// TIA Portal V20 program export: 0 tag tables, 53 data types, 23 data blocks, 177 code blocks (in call order from the OBs), 3 instance data blocks

TYPE "FRK_Access"
// stored: IsFailsafeCompliant false
   STRUCT
      CurrentLevel : DInt;
      CurrentUser : String[32];
      LoginFailed : Bool;
      Policy { S7_SetPoint := 'True'} : "ST_AccessPolicy";
      SessionGeneration : UDInt;
      LoginBusy : Bool;
      LoginResultSequence : UDInt;
      LoginTimeoutMs : UDInt;
      PolicySlot { ExternalAccessible := 'False'; ExternalVisible := 'False'; ExternalWritable := 'False'} : Int;
      PolicyLost { ExternalAccessible := 'False'; ExternalVisible := 'False'; ExternalWritable := 'False'} : Bool;
      PolicyLossAlarm { ExternalAccessible := 'False'; ExternalVisible := 'False'; ExternalWritable := 'False'} : Int;
      UserLossAlarm { ExternalAccessible := 'False'; ExternalVisible := 'False'; ExternalWritable := 'False'} : Int;
      ProviderGeneration { ExternalAccessible := 'False'; ExternalVisible := 'False'; ExternalWritable := 'False'} : UDInt;
      CandidateGeneration { ExternalAccessible := 'False'; ExternalVisible := 'False'; ExternalWritable := 'False'} : UDInt;
      ProviderEnabled { ExternalAccessible := 'False'; ExternalVisible := 'False'; ExternalWritable := 'False'} : Bool;
      LastActivity { ExternalAccessible := 'False'; ExternalVisible := 'False'; ExternalWritable := 'False'} : UDInt;
      LoginSince { ExternalAccessible := 'False'; ExternalVisible := 'False'; ExternalWritable := 'False'} : UDInt;
      LoginSequence { ExternalAccessible := 'False'; ExternalVisible := 'False'; ExternalWritable := 'False'} : UDInt;
      CandidateUser { ExternalAccessible := 'False'; ExternalVisible := 'False'; ExternalWritable := 'False'} : String[32];
      CandidateLevel { ExternalAccessible := 'False'; ExternalVisible := 'False'; ExternalWritable := 'False'} : DInt;
      Round { ExternalAccessible := 'False'; ExternalVisible := 'False'; ExternalWritable := 'False'} : DInt;
      Salt { ExternalAccessible := 'False'; ExternalVisible := 'False'; ExternalWritable := 'False'} : Array[0..15] of Byte;
      Digest { ExternalAccessible := 'False'; ExternalVisible := 'False'; ExternalWritable := 'False'} : Array[0..31] of Byte;
      Expected { ExternalAccessible := 'False'; ExternalVisible := 'False'; ExternalWritable := 'False'} : Array[0..31] of Byte;
   END_STRUCT;
END_TYPE

TYPE "FRK_AccessPolicyImage"
// stored: IsFailsafeCompliant false
   STRUCT
      SchemaVersion { ExternalAccessible := 'False'; ExternalVisible := 'False'; ExternalWritable := 'False'} : UInt;
      Scope { ExternalAccessible := 'False'; ExternalVisible := 'False'; ExternalWritable := 'False'} : String[80];
      Generation { ExternalAccessible := 'False'; ExternalVisible := 'False'; ExternalWritable := 'False'} : UDInt;
      Policy { ExternalAccessible := 'False'; ExternalVisible := 'False'; ExternalWritable := 'False'; S7_SetPoint := 'True'} : "ST_AccessPolicy";
      Checksum { ExternalAccessible := 'False'; ExternalVisible := 'False'; ExternalWritable := 'False'} : DWord;
   END_STRUCT;
END_TYPE

TYPE "FRK_AlarmLog"
// stored: IsFailsafeCompliant false
   STRUCT
      Active { S7_SetPoint := 'True'} : Array[1..16] of "ST_AlarmEvent";
      NActive : Int;
      Ring { S7_SetPoint := 'True'} : Array[1..64] of "ST_AlarmEvent";
      RingHead : Int;
      Blocking : Bool;
      Truncated : Bool;
      ComeMs { ExternalAccessible := 'False'; ExternalVisible := 'False'; ExternalWritable := 'False'} : Array[1..16] of UDInt;
      Automatic { ExternalAccessible := 'False'; ExternalVisible := 'False'; ExternalWritable := 'False'} : Array[1..16] of Bool;
      Touched { ExternalAccessible := 'False'; ExternalVisible := 'False'; ExternalWritable := 'False'} : Array[1..16] of Bool;
      RingUsed { ExternalAccessible := 'False'; ExternalVisible := 'False'; ExternalWritable := 'False'} : Int;
      SinkEnabled { ExternalAccessible := 'False'; ExternalVisible := 'False'; ExternalWritable := 'False'} : Bool;
   END_STRUCT;
END_TYPE

TYPE "FRK_Carrier"
// stored: IsFailsafeCompliant false
   STRUCT
      Enabled { ExternalAccessible := 'False'; ExternalVisible := 'False'; ExternalWritable := 'False'} : Bool;
      Kind { ExternalAccessible := 'False'; ExternalVisible := 'False'; ExternalWritable := 'False'} : DInt;
      Serial { ExternalAccessible := 'False'; ExternalVisible := 'False'; ExternalWritable := 'False'} : UDInt;
      Context { ExternalAccessible := 'False'; ExternalVisible := 'False'; ExternalWritable := 'False'; S7_SetPoint := 'True'} : "ST_PartContext";
      Written { ExternalAccessible := 'False'; ExternalVisible := 'False'; ExternalWritable := 'False'; S7_SetPoint := 'True'} : "ST_PartContext";
      Writes { ExternalAccessible := 'False'; ExternalVisible := 'False'; ExternalWritable := 'False'} : UDInt;
   END_STRUCT;
END_TYPE

TYPE "FRK_ConfigCursor"
// stored: IsFailsafeCompliant false
   STRUCT
      Position { ExternalAccessible := 'False'; ExternalVisible := 'False'; ExternalWritable := 'False'} : DInt;
      First { ExternalAccessible := 'False'; ExternalVisible := 'False'; ExternalWritable := 'False'} : DInt;
   END_STRUCT;
END_TYPE

TYPE "FRK_ConfigSlot"
// stored: IsFailsafeCompliant false
   STRUCT
      SchemaVersion { ExternalAccessible := 'False'; ExternalVisible := 'False'; ExternalWritable := 'False'} : UInt;
      Used { ExternalAccessible := 'False'; ExternalVisible := 'False'; ExternalWritable := 'False'} : Bool;
      ModelCode { ExternalAccessible := 'False'; ExternalVisible := 'False'; ExternalWritable := 'False'} : String[64];
      Record { ExternalAccessible := 'False'; ExternalVisible := 'False'; ExternalWritable := 'False'; S7_SetPoint := 'True'} : "ST_ConfigRecord";
   END_STRUCT;
END_TYPE

TYPE "FRK_ConfigValue"
// stored: IsFailsafeCompliant false
   STRUCT
      Number { ExternalAccessible := 'False'; ExternalVisible := 'False'; ExternalWritable := 'False'} : LInt;
      Flag { ExternalAccessible := 'False'; ExternalVisible := 'False'; ExternalWritable := 'False'} : Bool;
      Text { ExternalAccessible := 'False'; ExternalVisible := 'False'; ExternalWritable := 'False'} : String[80];
   END_STRUCT;
END_TYPE

TYPE "FRK_Core"
// stored: IsFailsafeCompliant false
   STRUCT
      Named { ExternalAccessible := 'False'; ExternalVisible := 'False'; ExternalWritable := 'False'} : Bool;
      Initialized { ExternalAccessible := 'False'; ExternalVisible := 'False'; ExternalWritable := 'False'} : Bool;
      RegIndex { ExternalAccessible := 'False'; ExternalVisible := 'False'; ExternalWritable := 'False'} : DInt;
      ParentIndex { ExternalAccessible := 'False'; ExternalVisible := 'False'; ExternalWritable := 'False'} : DInt;
      ModuleType { ExternalAccessible := 'False'; ExternalVisible := 'False'; ExternalWritable := 'False'} : DInt;
      Exec { ExternalAccessible := 'False'; ExternalVisible := 'False'; ExternalWritable := 'False'} : DInt;
      ExecPrev { ExternalAccessible := 'False'; ExternalVisible := 'False'; ExternalWritable := 'False'} : Bool;
      AbortPrev { ExternalAccessible := 'False'; ExternalVisible := 'False'; ExternalWritable := 'False'} : Bool;
      Armed { ExternalAccessible := 'False'; ExternalVisible := 'False'; ExternalWritable := 'False'} : Bool;
      Command { ExternalAccessible := 'False'; ExternalVisible := 'False'; ExternalWritable := 'False'} : DInt;
      CommandLabel { ExternalAccessible := 'False'; ExternalVisible := 'False'; ExternalWritable := 'False'} : String[120];
      Dispatch { ExternalAccessible := 'False'; ExternalVisible := 'False'; ExternalWritable := 'False'} : Bool;
      EvInit { ExternalAccessible := 'False'; ExternalVisible := 'False'; ExternalWritable := 'False'} : Bool;
      EvCommandStart { ExternalAccessible := 'False'; ExternalVisible := 'False'; ExternalWritable := 'False'} : Bool;
      ReleasePending { ExternalAccessible := 'False'; ExternalVisible := 'False'; ExternalWritable := 'False'} : Bool;
      EvAbort { ExternalAccessible := 'False'; ExternalVisible := 'False'; ExternalWritable := 'False'} : Bool;
      EvAbortInError { ExternalAccessible := 'False'; ExternalVisible := 'False'; ExternalWritable := 'False'} : Bool;
      EvModeExit { ExternalAccessible := 'False'; ExternalVisible := 'False'; ExternalWritable := 'False'} : Bool;
      EvModeChanged { ExternalAccessible := 'False'; ExternalVisible := 'False'; ExternalWritable := 'False'} : Bool;
      "Step" { ExternalAccessible := 'False'; ExternalVisible := 'False'; ExternalWritable := 'False'} : DInt;
      HookResult { ExternalAccessible := 'False'; ExternalVisible := 'False'; ExternalWritable := 'False'} : DInt;
      Held { ExternalAccessible := 'False'; ExternalVisible := 'False'; ExternalWritable := 'False'} : Bool;
      HoldReq { ExternalAccessible := 'False'; ExternalVisible := 'False'; ExternalWritable := 'False'} : Bool;
      HoldReason { ExternalAccessible := 'False'; ExternalVisible := 'False'; ExternalWritable := 'False'} : DInt;
      DiagTouched { ExternalAccessible := 'False'; ExternalVisible := 'False'; ExternalWritable := 'False'} : Bool;
      TimingOpen { ExternalAccessible := 'False'; ExternalVisible := 'False'; ExternalWritable := 'False'} : Bool;
      StartMs { ExternalAccessible := 'False'; ExternalVisible := 'False'; ExternalWritable := 'False'} : UDInt;
      LastNowMs { ExternalAccessible := 'False'; ExternalVisible := 'False'; ExternalWritable := 'False'} : UDInt;
      DeltaMs { ExternalAccessible := 'False'; ExternalVisible := 'False'; ExternalWritable := 'False'} : UDInt;
      ActiveMs { ExternalAccessible := 'False'; ExternalVisible := 'False'; ExternalWritable := 'False'} : UDInt;
      TimeoutMs { ExternalAccessible := 'False'; ExternalVisible := 'False'; ExternalWritable := 'False'} : UDInt;
      Timing { ExternalAccessible := 'False'; ExternalVisible := 'False'; ExternalWritable := 'False'; S7_SetPoint := 'True'} : "ST_ModuleTiming";
      FaultSlot { ExternalAccessible := 'False'; ExternalVisible := 'False'; ExternalWritable := 'False'} : Int;
      FaultHandled { ExternalAccessible := 'False'; ExternalVisible := 'False'; ExternalWritable := 'False'} : Bool;
   END_STRUCT;
END_TYPE

TYPE "FRK_DecisionSlot"
// stored: IsFailsafeCompliant false
   STRUCT
      RootIndex { ExternalAccessible := 'False'; ExternalVisible := 'False'; ExternalWritable := 'False'} : DInt;
      Owner { ExternalAccessible := 'False'; ExternalVisible := 'False'; ExternalWritable := 'False'} : DInt;
      Request { ExternalAccessible := 'False'; ExternalVisible := 'False'; ExternalWritable := 'False'; S7_SetPoint := 'True'} : "ST_DecisionRequest";
      Answer { ExternalAccessible := 'False'; ExternalVisible := 'False'; ExternalWritable := 'False'} : Int;
      AskedAt { ExternalAccessible := 'False'; ExternalVisible := 'False'; ExternalWritable := 'False'} : UDInt;
      OverlapLogged { ExternalAccessible := 'False'; ExternalVisible := 'False'; ExternalWritable := 'False'} : Bool;
      ResolutionLogged { ExternalAccessible := 'False'; ExternalVisible := 'False'; ExternalWritable := 'False'} : Bool;
   END_STRUCT;
END_TYPE

TYPE "FRK_JsonField"
// stored: IsFailsafeCompliant false
   STRUCT
      Key { ExternalAccessible := 'False'; ExternalVisible := 'False'; ExternalWritable := 'False'} : String[16];
      Text { ExternalAccessible := 'False'; ExternalVisible := 'False'; ExternalWritable := 'False'} : WString[160];
      Quoted { ExternalAccessible := 'False'; ExternalVisible := 'False'; ExternalWritable := 'False'} : Bool;
   END_STRUCT;
END_TYPE

TYPE "FRK_ManualConditionRow"
// stored: IsFailsafeCompliant false
   STRUCT
      Used { ExternalAccessible := 'False'; ExternalVisible := 'False'; ExternalWritable := 'False'} : Bool;
      Value { ExternalAccessible := 'False'; ExternalVisible := 'False'; ExternalWritable := 'False'} : DInt;
      Ok { ExternalAccessible := 'False'; ExternalVisible := 'False'; ExternalWritable := 'False'} : Bool;
      Diag { ExternalAccessible := 'False'; ExternalVisible := 'False'; ExternalWritable := 'False'; S7_SetPoint := 'True'} : "ST_Diagnostic";
      Bypassable { ExternalAccessible := 'False'; ExternalVisible := 'False'; ExternalWritable := 'False'} : Bool;
   END_STRUCT;
END_TYPE

TYPE "FRK_RegistryRow"
// stored: IsFailsafeCompliant false
   STRUCT
      Valid { ExternalAccessible := 'False'; ExternalVisible := 'False'; ExternalWritable := 'False'} : Bool;
      Parent { ExternalAccessible := 'False'; ExternalVisible := 'False'; ExternalWritable := 'False'} : DInt;
      ModuleType { ExternalAccessible := 'False'; ExternalVisible := 'False'; ExternalWritable := 'False'} : DInt;
      TypeId { ExternalAccessible := 'False'; ExternalVisible := 'False'; ExternalWritable := 'False'} : DInt;
      Capabilities { ExternalAccessible := 'False'; ExternalVisible := 'False'; ExternalWritable := 'False'} : DWord;
      Exec { ExternalAccessible := 'False'; ExternalVisible := 'False'; ExternalWritable := 'False'} : DInt;
      ReasonCode { ExternalAccessible := 'False'; ExternalVisible := 'False'; ExternalWritable := 'False'} : DInt;
      Severity { ExternalAccessible := 'False'; ExternalVisible := 'False'; ExternalWritable := 'False'} : DInt;
      AlarmBlocking { ExternalAccessible := 'False'; ExternalVisible := 'False'; ExternalWritable := 'False'} : Bool;
   END_STRUCT;
END_TYPE

TYPE "FRK_SetPayload"
// stored: IsFailsafeCompliant false
   STRUCT
      Info { ExternalAccessible := 'False'; ExternalVisible := 'False'; ExternalWritable := 'False'; S7_SetPoint := 'True'} : "ST_ConfigSetInfo";
      Records { ExternalAccessible := 'False'; ExternalVisible := 'False'; ExternalWritable := 'False'; S7_SetPoint := 'True'} : Array[1..24] of "ST_ConfigRecord";
   END_STRUCT;
END_TYPE

TYPE "FRK_SetWorkspace"
// stored: IsFailsafeCompliant false
   STRUCT
      Payload { ExternalAccessible := 'False'; ExternalVisible := 'False'; ExternalWritable := 'False'; S7_SetPoint := 'True'} : "FRK_SetPayload";
      Seen { ExternalAccessible := 'False'; ExternalVisible := 'False'; ExternalWritable := 'False'} : Array[1..24] of Bool;
      Matched { ExternalAccessible := 'False'; ExternalVisible := 'False'; ExternalWritable := 'False'} : Int;
      RejectScope { ExternalAccessible := 'False'; ExternalVisible := 'False'; ExternalWritable := 'False'} : String[80];
      RejectKey { ExternalAccessible := 'False'; ExternalVisible := 'False'; ExternalWritable := 'False'} : String[160];
      Importing { ExternalAccessible := 'False'; ExternalVisible := 'False'; ExternalWritable := 'False'} : Bool;
      Exporting { ExternalAccessible := 'False'; ExternalVisible := 'False'; ExternalWritable := 'False'} : Bool;
      NextLine { ExternalAccessible := 'False'; ExternalVisible := 'False'; ExternalWritable := 'False'} : Int;
      Generation { ExternalAccessible := 'False'; ExternalVisible := 'False'; ExternalWritable := 'False'} : UDInt;
      Received { ExternalAccessible := 'False'; ExternalVisible := 'False'; ExternalWritable := 'False'} : Int;
      Piece { ExternalAccessible := 'False'; ExternalVisible := 'False'; ExternalWritable := 'False'} : WString[480];
      Line { ExternalAccessible := 'False'; ExternalVisible := 'False'; ExternalWritable := 'False'} : WString[480];
      Fields { ExternalAccessible := 'False'; ExternalVisible := 'False'; ExternalWritable := 'False'; S7_SetPoint := 'True'} : Array[1..9] of "FRK_JsonField";
      FieldCount { ExternalAccessible := 'False'; ExternalVisible := 'False'; ExternalWritable := 'False'} : Int;
   END_STRUCT;
END_TYPE

TYPE "FRK_Unit"
// stored: IsFailsafeCompliant false
   STRUCT
      Initialized { ExternalAccessible := 'False'; ExternalVisible := 'False'; ExternalWritable := 'False'} : Bool;
      Mode { ExternalAccessible := 'False'; ExternalVisible := 'False'; ExternalWritable := 'False'} : DInt;
      RequestedMode { ExternalAccessible := 'False'; ExternalVisible := 'False'; ExternalWritable := 'False'} : DInt;
      ModePending { ExternalAccessible := 'False'; ExternalVisible := 'False'; ExternalWritable := 'False'} : Bool;
      ExitFirst { ExternalAccessible := 'False'; ExternalVisible := 'False'; ExternalWritable := 'False'} : Bool;
      RunReq { ExternalAccessible := 'False'; ExternalVisible := 'False'; ExternalWritable := 'False'} : Bool;
      AbortReq { ExternalAccessible := 'False'; ExternalVisible := 'False'; ExternalWritable := 'False'} : Bool;
      StopReq { ExternalAccessible := 'False'; ExternalVisible := 'False'; ExternalWritable := 'False'} : Bool;
      ModeSince { ExternalAccessible := 'False'; ExternalVisible := 'False'; ExternalWritable := 'False'} : UDInt;
      ReleaseChildren { ExternalAccessible := 'False'; ExternalVisible := 'False'; ExternalWritable := 'False'} : Bool;
      Clearing { ExternalAccessible := 'False'; ExternalVisible := 'False'; ExternalWritable := 'False'} : Bool;
      FaultLatched { ExternalAccessible := 'False'; ExternalVisible := 'False'; ExternalWritable := 'False'} : Bool;
      PrevError { ExternalAccessible := 'False'; ExternalVisible := 'False'; ExternalWritable := 'False'} : Bool;
      EvReset { ExternalAccessible := 'False'; ExternalVisible := 'False'; ExternalWritable := 'False'} : Bool;
      SeenSequence { ExternalAccessible := 'False'; ExternalVisible := 'False'; ExternalWritable := 'False'} : UDInt;
      RequestPending { ExternalAccessible := 'False'; ExternalVisible := 'False'; ExternalWritable := 'False'} : Bool;
      Request { ExternalAccessible := 'False'; ExternalVisible := 'False'; ExternalWritable := 'False'; S7_SetPoint := 'True'} : "ST_HmiRequest";
      RequestUser { ExternalAccessible := 'False'; ExternalVisible := 'False'; ExternalWritable := 'False'} : String[32];
      Permit { ExternalAccessible := 'False'; ExternalVisible := 'False'; ExternalWritable := 'False'} : Bool;
      PermitDiag { ExternalAccessible := 'False'; ExternalVisible := 'False'; ExternalWritable := 'False'; S7_SetPoint := 'True'} : "ST_Diagnostic";
      CarrierIndex { ExternalAccessible := 'False'; ExternalVisible := 'False'; ExternalWritable := 'False'} : DInt;
      Good { ExternalAccessible := 'False'; ExternalVisible := 'False'; ExternalWritable := 'False'} : UDInt;
      Nok { ExternalAccessible := 'False'; ExternalVisible := 'False'; ExternalWritable := 'False'} : UDInt;
      Rework { ExternalAccessible := 'False'; ExternalVisible := 'False'; ExternalWritable := 'False'} : UDInt;
      NokReason { ExternalAccessible := 'False'; ExternalVisible := 'False'; ExternalWritable := 'False'} : DInt;
      CascadePending { ExternalAccessible := 'False'; ExternalVisible := 'False'; ExternalWritable := 'False'} : Bool;
      CascadeKind { ExternalAccessible := 'False'; ExternalVisible := 'False'; ExternalWritable := 'False'} : DInt;
      CascadeMode { ExternalAccessible := 'False'; ExternalVisible := 'False'; ExternalWritable := 'False'} : DInt;
      FollowStart { ExternalAccessible := 'False'; ExternalVisible := 'False'; ExternalWritable := 'False'} : Bool;
      AlarmBlocking { ExternalAccessible := 'False'; ExternalVisible := 'False'; ExternalWritable := 'False'} : Bool;
      ConfigBlocked { ExternalAccessible := 'False'; ExternalVisible := 'False'; ExternalWritable := 'False'} : Bool;
      ConfigEnabled { ExternalAccessible := 'False'; ExternalVisible := 'False'; ExternalWritable := 'False'} : Bool;
      ModelEnabled { ExternalAccessible := 'False'; ExternalVisible := 'False'; ExternalWritable := 'False'} : Bool;
      ConfigSetsEnabled { ExternalAccessible := 'False'; ExternalVisible := 'False'; ExternalWritable := 'False'} : Bool;
   END_STRUCT;
END_TYPE

TYPE "ST_AccessPolicy"
// stored: IsFailsafeCompliant false
   STRUCT
      Required : Array[0..11] of DInt;
      SessionTimeout : Time := T#0MS;
   END_STRUCT;
END_TYPE

TYPE "ST_AlarmEvent"
// stored: IsFailsafeCompliant false
   STRUCT
      ReasonCode : DInt;
      Description : WString[255];
      SourcePath : WString[255];
      IoTag : String[80];
      IoAddress : String[80];
      Severity : DInt;
      Category : DInt;
      ResetClass : DInt;
      State : DInt;
      ComeAt : LDT;
      GoneAt : LDT;
      ResetAt : LDT;
      Duration : Time;
      Shelved : Bool;
      ShelvedUntil : LDT;
      ComeTimeSynchronized : Bool;
      GoneTimeSynchronized : Bool;
      ResetTimeSynchronized : Bool;
      ShelfTimeSynchronized : Bool;
   END_STRUCT;
END_TYPE

TYPE "ST_CommandInfo"
// stored: IsFailsafeCompliant false
   STRUCT
      Value : DInt;
      Label : String[120];
      Style : DInt;
   END_STRUCT;
END_TYPE

TYPE "ST_ConfigEntry"
// stored: IsFailsafeCompliant false
   STRUCT
      Scope : WString[255];
      Item : WString[255];
      ValueText : WString[255];
      WriteKey : String[160];
      WriteRevision : UDInt;
      ConfigKind : DInt;
      ValueType : DInt;
      Writable : Bool;
      RequiresReady : Bool;
      HasMinimum : Bool;
      HasMaximum : Bool;
      Minimum : LReal;
      Maximum : LReal;
      Unit : String[16];
      LabelKey : String[160];
      EnumDomain : WString[255];
      ClassId : String[40];
      ReadLevel : DInt;
      WriteLevel : DInt;
      Readable : Bool;
      UnitCode : DInt;
      EnumLabelKey : String[80];
      ModelScoped : Bool;
   END_STRUCT;
END_TYPE

TYPE "ST_ConfigPage"
// stored: IsFailsafeCompliant false
   STRUCT
      Revision : UDInt;
      PageIndex : Int;
      PageCount : Int;
      EntryCount : Int;
      Entries { S7_SetPoint := 'True'} : Array[1..16] of "ST_ConfigEntry";
   END_STRUCT;
END_TYPE

TYPE "ST_ConfigPersistStatus"
// stored: IsFailsafeCompliant false
   STRUCT
      Pending : Bool;
      Failed : Bool;
      WindowMs : UDInt := 5000;
      PendingSince : LDT;
      StorePresent : Bool;
      StoreKind : DInt;
      RestorePolicy : DInt;
      RestoreLost : Bool;
      RestoreAcknowledged : Bool;
      LostPath : String[80];
      LastSetName : String[80];
      LastSetRecords : Int;
      LastRejectScope : String[80];
      LastRejectKey : String[160];
   END_STRUCT;
END_TYPE

TYPE "ST_ConfigRecord"
// stored: IsFailsafeCompliant false
   STRUCT
      Scope : String[80];
      WriteKey : String[160];
      Revision : UDInt;
      Kind : DInt;
      ValueType : DInt;
      ValueText : String[80];
   END_STRUCT;
END_TYPE

TYPE "ST_ConfigSetInfo"
// stored: IsFailsafeCompliant false
   STRUCT
      Used : Bool;
      SetName : String[80];
      RootIdentity : String[80];
      SetSchema : UInt;
      ConfigRev : UDInt;
      Kind : DInt;
      ModelCode : String[64];
      RecordCount : Int;
      CreatedAt : LDT;
      TimeSynchronized : Bool;
   END_STRUCT;
END_TYPE

TYPE "ST_DecisionRequest"
// stored: IsFailsafeCompliant false
   STRUCT
      Prompt : WString[255];
      Options : Array[1..6] of String[64];
      Default : Int;
      Timeout : Time;
      SourcePath : WString[255];
   END_STRUCT;
END_TYPE

TYPE "ST_DeclarationCellHal"
// stored: IsFailsafeCompliant false
   STRUCT
      Clamp { ExternalAccessible := 'False'; ExternalVisible := 'False'; ExternalWritable := 'False'; S7_SetPoint := 'True'} : "ST_DeclarationLeafHal";
      Gate { ExternalAccessible := 'False'; ExternalVisible := 'False'; ExternalWritable := 'False'; S7_SetPoint := 'True'} : "ST_DeclarationLeafHal";
   END_STRUCT;
END_TYPE

TYPE "ST_DeclarationLeafHal"
// stored: IsFailsafeCompliant false
   STRUCT
      Sample : DInt;
      Permit : Bool := TRUE;
      Finish : Bool;
      BackgroundFault : Bool;
      Diag { S7_SetPoint := 'True'} : "ST_Diagnostic";
      LaterDiag { S7_SetPoint := 'True'} : "ST_Diagnostic";
      ExitHold : Bool;
      Verdict : DInt := 1;
   END_STRUCT;
END_TYPE

TYPE "ST_DeclarationOutCmd"
// stored: IsFailsafeCompliant false
   STRUCT
      Result : DInt;
   END_STRUCT;
END_TYPE

TYPE "ST_DeclarationOutImm"
// stored: IsFailsafeCompliant false
   STRUCT
      Sample : DInt;
      InitCount : DInt;
      StartCount : DInt;
      CyclicCount : DInt;
      AbortCount : DInt;
      ErrorAbortCount : DInt;
      DispatchCount : DInt;
      SeenValue : DInt;
      Ordered : Bool;
      Output : Bool;
   END_STRUCT;
END_TYPE

TYPE "ST_DeclarationParCfg"
// stored: IsFailsafeCompliant false
   STRUCT
      SchemaVersion : UInt := 4;
      Timeout : Time := T#8S;
      Preset : DInt := 10;
   END_STRUCT;
END_TYPE

TYPE "ST_DeclarationParCmd"
// stored: IsFailsafeCompliant false
   STRUCT
      Value : DInt;
   END_STRUCT;
END_TYPE

TYPE "ST_DeclarationUnitHal"
// stored: IsFailsafeCompliant false
   STRUCT
      Cell { ExternalAccessible := 'False'; ExternalVisible := 'False'; ExternalWritable := 'False'; S7_SetPoint := 'True'} : "ST_DeclarationCellHal";
      Satellite { ExternalAccessible := 'False'; ExternalVisible := 'False'; ExternalWritable := 'False'; S7_SetPoint := 'True'} : "ST_SatelliteUnitHal";
   END_STRUCT;
END_TYPE

TYPE "ST_Diagnostic"
// stored: IsFailsafeCompliant false
   STRUCT
      ReasonCode : DInt;
      SourcePath : WString[255];
      Description : WString[255];
      IoTag : String[80];
      IoAddress : String[80];
      Severity : DInt;
      Category : DInt;
      Since : LDT;
      TimeSynchronized : Bool;
   END_STRUCT;
END_TYPE

TYPE "ST_FraktalHal"
// stored: IsFailsafeCompliant false
   STRUCT
      StationA { ExternalAccessible := 'False'; ExternalVisible := 'False'; ExternalWritable := 'False'; S7_SetPoint := 'True'} : "ST_DeclarationUnitHal";
      StationB { ExternalAccessible := 'False'; ExternalVisible := 'False'; ExternalWritable := 'False'; S7_SetPoint := 'True'} : "ST_DeclarationUnitHal";
   END_STRUCT;
END_TYPE

TYPE "ST_HmiRequest"
// stored: IsFailsafeCompliant false
   STRUCT
      Kind : DInt;
      TargetPath : WString[255];
      NameValue : String[160];
      TextValue : WString[255];
      User : String[32];
      Secret : String[32];
      IntValue : DInt;
      BoolValue : Bool;
      DurationMs : UDInt;
      Sequence : UDInt;
   END_STRUCT;
END_TYPE

TYPE "ST_HmiResponse"
// stored: IsFailsafeCompliant false
   STRUCT
      AckSequence : UDInt;
      Accepted : Bool;
      Diagnostic : WString[255];
      Report { S7_SetPoint := 'True'} : "ST_ReleaseReport";
      ConfigPage { S7_SetPoint := 'True'} : "ST_ConfigPage";
   END_STRUCT;
END_TYPE

TYPE "ST_InnerUnitHal"
// stored: IsFailsafeCompliant false
   STRUCT
      Cell { ExternalAccessible := 'False'; ExternalVisible := 'False'; ExternalWritable := 'False'; S7_SetPoint := 'True'} : "ST_DeclarationCellHal";
   END_STRUCT;
END_TYPE

TYPE "ST_MeasRecord"
// stored: IsFailsafeCompliant false
   STRUCT
      "Name" : String[64];
      Value : LReal;
      Minimum : LReal;
      Maximum : LReal;
      Target : LReal;
      Unit : String[16];
      InTol : Bool;
   END_STRUCT;
END_TYPE

TYPE "ST_ModePolicy"
// stored: IsFailsafeCompliant false
   STRUCT
      Shield : DInt;
      Style : DInt;
   END_STRUCT;
END_TYPE

TYPE "ST_ModelField"
// stored: IsFailsafeCompliant false
   STRUCT
      "Name" : String[32];
      Value : String[64];
   END_STRUCT;
END_TYPE

TYPE "ST_ModelId"
// stored: IsFailsafeCompliant false
   STRUCT
      ModelCode : String[64];
      "Family" : String[64];
      Variant : String[64];
      Fields { S7_SetPoint := 'True'} : Array[1..8] of "ST_ModelField";
      NField : Int;
   END_STRUCT;
END_TYPE

TYPE "ST_ModuleStatus"
// stored: IsFailsafeCompliant false
   STRUCT
      "Name" : String[80];
      DisplayNameKey : String[160];
      DescriptionKey : String[160];
      TypeKey : String[160];
      ModuleType : DInt;
      State : DInt;
      FaultActive : Bool;
      Diagnostic { S7_SetPoint := 'True'} : "ST_Diagnostic";
      TileEnable : Bool := TRUE;
      ControlDomainId : String[80];
   END_STRUCT;
END_TYPE

TYPE "ST_ModuleTiming"
// stored: IsFailsafeCompliant false
   STRUCT
      LastCmdTime : Time;
      Rows { S7_SetPoint := 'True'} : Array[1..8] of "ST_TimingRow";
      Truncated : Bool;
   END_STRUCT;
END_TYPE

TYPE "ST_PartContext"
// stored: IsFailsafeCompliant false
   STRUCT
      Uid : String[64];
      Present : Bool;
      CarrierKind : DInt;
      Result { S7_SetPoint := 'True'} : "ST_PartResult";
      Parents : Array[1..8] of String[64];
   END_STRUCT;
END_TYPE

TYPE "ST_PartResult"
// stored: IsFailsafeCompliant false
   STRUCT
      Verdict : DInt;
      ReasonCode : DInt;
      Records { S7_SetPoint := 'True'} : Array[1..32] of "ST_MeasRecord";
      StationPath : WString[255];
      Stamp : LDT;
      TimeSynchronized : Bool;
   END_STRUCT;
END_TYPE

TYPE "ST_ReleaseReason"
// stored: IsFailsafeCompliant false
   STRUCT
      Description : WString[255];
      ReasonCode : DInt;
      SourcePath : WString[255];
      Kind : DInt;
      Bypassable : Bool;
   END_STRUCT;
END_TYPE

TYPE "ST_ReleaseReport"
// stored: IsFailsafeCompliant false
   STRUCT
      Released : Bool;
      Count : Int;
      Reasons { S7_SetPoint := 'True'} : Array[1..24] of "ST_ReleaseReason";
   END_STRUCT;
END_TYPE

TYPE "ST_SatelliteUnitHal"
// stored: IsFailsafeCompliant false
   STRUCT
      Cell { ExternalAccessible := 'False'; ExternalVisible := 'False'; ExternalWritable := 'False'; S7_SetPoint := 'True'} : "ST_DeclarationCellHal";
      Inner { ExternalAccessible := 'False'; ExternalVisible := 'False'; ExternalWritable := 'False'; S7_SetPoint := 'True'} : "ST_InnerUnitHal";
   END_STRUCT;
END_TYPE

TYPE "ST_StateFlag"
// stored: IsFailsafeCompliant false
   STRUCT
      Key : String[120];
      Value : Bool;
      Since : LDT;
      Stale : Bool;
   END_STRUCT;
END_TYPE

TYPE "ST_TimingRow"
// stored: IsFailsafeCompliant false
   STRUCT
      Id : DInt;
      Label : String[120];
      TimeClass : DInt;
      Count : UDInt;
      Last : Time;
      Minimum : Time;
      Maximum : Time;
      Avg : Time;
   END_STRUCT;
END_TYPE

TYPE "ST_UnitProbeDevice"
// stored: IsFailsafeCompliant false
   STRUCT
      Cycles : UDInt;
      ExitCalls : UDInt;
      Changes : UDInt;
      Resets : UDInt;
      Received : Bool;
      Processed : Bool;
   END_STRUCT;
END_TYPE

TYPE "ST_UnitProbeImm"
// stored: IsFailsafeCompliant false
   STRUCT
      Cycles : UDInt;
      ExitCalls : UDInt;
      Changes : UDInt;
      Resets : UDInt;
      AtHome : Bool;
   END_STRUCT;
END_TYPE

TYPE "ST_UnitProbeStationCfg"
// stored: IsFailsafeCompliant false
   STRUCT
      SchemaVersion : UInt := 2;
      SiteLabel : String[80] := 'bench';
      Enabled : Bool := TRUE;
      LongText : String[80] := 'long default';
   END_STRUCT;
END_TYPE

TYPE "ST_UserRecord"
// stored: IsFailsafeCompliant false
   STRUCT
      User : String[32];
      Salt : Array[0..15] of Byte;
      PinHash : Array[0..31] of Byte;
      Level : DInt;
   END_STRUCT;
END_TYPE

DATA_BLOCK "FRK_AccessPolicies"   // DB3
{ S7_Optimized_Access := 'TRUE' }
VERSION : 0.1
// stored: AutoNumber true, DBAccessibleFromOPCUA true, DBAccessibleFromWebserver true, IsOnlyStoredInLoadMemory false, IsRetainMemResEnabled false, IsWriteProtectedInAS false, MemoryReserve 100
   VAR RETAIN
      Rows { ExternalAccessible := 'False'; ExternalVisible := 'False'; ExternalWritable := 'False'; S7_SetPoint := 'True'} : Array[1..2] of "FRK_AccessPolicyImage";
   END_VAR
BEGIN
END_DATA_BLOCK

DATA_BLOCK "FRK_AccessStorage"   // DB4
{ S7_Optimized_Access := 'TRUE' }
VERSION : 0.1
// stored: AutoNumber true, DBAccessibleFromOPCUA true, DBAccessibleFromWebserver true, IsOnlyStoredInLoadMemory false, IsRetainMemResEnabled false, IsWriteProtectedInAS false, MemoryReserve 100
   VAR
      UsersReady { ExternalAccessible := 'False'; ExternalVisible := 'False'; ExternalWritable := 'False'} : Bool;
      UsersLost { ExternalAccessible := 'False'; ExternalVisible := 'False'; ExternalWritable := 'False'} : Bool;
      EmptyPolicy { ExternalAccessible := 'False'; ExternalVisible := 'False'; ExternalWritable := 'False'; S7_SetPoint := 'True'} : "ST_AccessPolicy";
   END_VAR
BEGIN
END_DATA_BLOCK

DATA_BLOCK "FRK_Carriers"   // DB5
{ S7_Optimized_Access := 'TRUE' }
VERSION : 0.1
// stored: AutoNumber true, DBAccessibleFromOPCUA true, DBAccessibleFromWebserver true, IsOnlyStoredInLoadMemory false, IsRetainMemResEnabled false, IsWriteProtectedInAS false, MemoryReserve 100
   VAR
      Slots { ExternalAccessible := 'False'; ExternalVisible := 'False'; ExternalWritable := 'False'; S7_SetPoint := 'True'} : Array[0..32] of "FRK_Carrier";
   END_VAR
BEGIN
END_DATA_BLOCK

DATA_BLOCK "FRK_Clock"   // DB1
{ S7_Optimized_Access := 'TRUE' }
VERSION : 0.1
// stored: AutoNumber true, DBAccessibleFromOPCUA true, DBAccessibleFromWebserver true, IsOnlyStoredInLoadMemory false, IsRetainMemResEnabled false, IsWriteProtectedInAS false, MemoryReserve 100
   VAR
      Mem { ExternalAccessible := 'False'; ExternalVisible := 'False'; ExternalWritable := 'False'} : LReal;
      AccMs { ExternalAccessible := 'False'; ExternalVisible := 'False'; ExternalWritable := 'False'} : LReal;
      NowMs { ExternalAccessible := 'False'; ExternalVisible := 'False'; ExternalWritable := 'False'} : UDInt;
   END_VAR
BEGIN
END_DATA_BLOCK

DATA_BLOCK "FRK_ConfigRuntime"   // DB6
{ S7_Optimized_Access := 'TRUE' }
VERSION : 0.1
// stored: AutoNumber true, DBAccessibleFromOPCUA true, DBAccessibleFromWebserver true, IsOnlyStoredInLoadMemory false, IsRetainMemResEnabled false, IsWriteProtectedInAS false, MemoryReserve 100
   VAR
      Fresh { ExternalAccessible := 'False'; ExternalVisible := 'False'; ExternalWritable := 'False'} : Bool;
      Unavailable { ExternalAccessible := 'False'; ExternalVisible := 'False'; ExternalWritable := 'False'} : Bool;
      Failed { ExternalAccessible := 'False'; ExternalVisible := 'False'; ExternalWritable := 'False'} : Array[1..2] of Bool;
      LossSlot { ExternalAccessible := 'False'; ExternalVisible := 'False'; ExternalWritable := 'False'} : Array[1..2] of Int;
   END_VAR
BEGIN
END_DATA_BLOCK

DATA_BLOCK "FRK_ConfigScratch"   // DB7
{ S7_Optimized_Access := 'TRUE' }
VERSION : 0.1
// stored: AutoNumber true, DBAccessibleFromOPCUA true, DBAccessibleFromWebserver true, IsOnlyStoredInLoadMemory false, IsRetainMemResEnabled false, IsWriteProtectedInAS false, MemoryReserve 100
   VAR
      Entry { ExternalAccessible := 'False'; ExternalVisible := 'False'; ExternalWritable := 'False'; S7_SetPoint := 'True'} : "ST_ConfigEntry";
      Blank { ExternalAccessible := 'False'; ExternalVisible := 'False'; ExternalWritable := 'False'; S7_SetPoint := 'True'} : "ST_ConfigEntry";
      Value { ExternalAccessible := 'False'; ExternalVisible := 'False'; ExternalWritable := 'False'; S7_SetPoint := 'True'} : "FRK_ConfigValue";
      Storage { ExternalAccessible := 'False'; ExternalVisible := 'False'; ExternalWritable := 'False'} : DInt;
      Schema { ExternalAccessible := 'False'; ExternalVisible := 'False'; ExternalWritable := 'False'} : UInt;
      Minimum { ExternalAccessible := 'False'; ExternalVisible := 'False'; ExternalWritable := 'False'} : LReal;
      Maximum { ExternalAccessible := 'False'; ExternalVisible := 'False'; ExternalWritable := 'False'} : LReal;
      MaxLength { ExternalAccessible := 'False'; ExternalVisible := 'False'; ExternalWritable := 'False'} : Int;
      MinRead { ExternalAccessible := 'False'; ExternalVisible := 'False'; ExternalWritable := 'False'} : DInt;
      MinWrite { ExternalAccessible := 'False'; ExternalVisible := 'False'; ExternalWritable := 'False'} : DInt;
   END_VAR
BEGIN
END_DATA_BLOCK

DATA_BLOCK "FRK_ConfigStore"   // DB8
{ S7_Optimized_Access := 'TRUE' }
VERSION : 0.1
// stored: AutoNumber true, DBAccessibleFromOPCUA true, DBAccessibleFromWebserver true, IsOnlyStoredInLoadMemory false, IsRetainMemResEnabled false, IsWriteProtectedInAS false, MemoryReserve 100
   VAR RETAIN
      SchemaVersion { ExternalAccessible := 'False'; ExternalVisible := 'False'; ExternalWritable := 'False'} : UInt;
      Rows { ExternalAccessible := 'False'; ExternalVisible := 'False'; ExternalWritable := 'False'; S7_SetPoint := 'True'} : Array[1..114] of "FRK_ConfigSlot";
      ActiveModels { ExternalAccessible := 'False'; ExternalVisible := 'False'; ExternalWritable := 'False'} : Array[1..2] of String[64];
      Lost { ExternalAccessible := 'False'; ExternalVisible := 'False'; ExternalWritable := 'False'} : Array[1..2] of Bool;
      Acknowledged { ExternalAccessible := 'False'; ExternalVisible := 'False'; ExternalWritable := 'False'} : Array[1..2] of Bool;
      LostPath { ExternalAccessible := 'False'; ExternalVisible := 'False'; ExternalWritable := 'False'} : Array[1..2] of String[80];
   END_VAR
BEGIN
END_DATA_BLOCK

DATA_BLOCK "FRK_Decisions"   // DB9
{ S7_Optimized_Access := 'TRUE' }
VERSION : 0.1
// stored: AutoNumber true, DBAccessibleFromOPCUA true, DBAccessibleFromWebserver true, IsOnlyStoredInLoadMemory false, IsRetainMemResEnabled false, IsWriteProtectedInAS false, MemoryReserve 100
   VAR
      Slots { ExternalAccessible := 'False'; ExternalVisible := 'False'; ExternalWritable := 'False'; S7_SetPoint := 'True'} : Array[1..2] of "FRK_DecisionSlot";
      EmptyRequest { ExternalAccessible := 'False'; ExternalVisible := 'False'; ExternalWritable := 'False'; S7_SetPoint := 'True'} : "ST_DecisionRequest";
   END_VAR
BEGIN
END_DATA_BLOCK

DATA_BLOCK "FRK_LocalUsers"   // DB10
{ S7_Optimized_Access := 'TRUE' }
VERSION : 0.1
// stored: AutoNumber true, DBAccessibleFromOPCUA true, DBAccessibleFromWebserver true, IsOnlyStoredInLoadMemory false, IsRetainMemResEnabled false, IsWriteProtectedInAS false, MemoryReserve 100
   VAR RETAIN
      SchemaVersion { ExternalAccessible := 'False'; ExternalVisible := 'False'; ExternalWritable := 'False'} : UInt;
      Generation { ExternalAccessible := 'False'; ExternalVisible := 'False'; ExternalWritable := 'False'} : UDInt;
      Count { ExternalAccessible := 'False'; ExternalVisible := 'False'; ExternalWritable := 'False'} : DInt;
      Rows { ExternalAccessible := 'False'; ExternalVisible := 'False'; ExternalWritable := 'False'; S7_SetPoint := 'True'} : Array[1..16] of "ST_UserRecord";
      Checksum { ExternalAccessible := 'False'; ExternalVisible := 'False'; ExternalWritable := 'False'} : DWord;
   END_VAR
BEGIN
END_DATA_BLOCK

DATA_BLOCK "FRK_Registry"   // DB2
{ S7_Optimized_Access := 'TRUE' }
VERSION : 0.1
// stored: AutoNumber true, DBAccessibleFromOPCUA true, DBAccessibleFromWebserver true, IsOnlyStoredInLoadMemory false, IsRetainMemResEnabled false, IsWriteProtectedInAS false, MemoryReserve 100
   VAR
      Count { ExternalAccessible := 'False'; ExternalVisible := 'False'; ExternalWritable := 'False'} : DInt;
      Fault { ExternalAccessible := 'False'; ExternalVisible := 'False'; ExternalWritable := 'False'} : Bool;
      Rows { ExternalAccessible := 'False'; ExternalVisible := 'False'; ExternalWritable := 'False'; S7_SetPoint := 'True'} : Array[0..32] of "FRK_RegistryRow";
   END_VAR
BEGIN
END_DATA_BLOCK

DATA_BLOCK "FRK_SetRuntime"   // DB11
{ S7_Optimized_Access := 'TRUE' }
VERSION : 0.1
// stored: AutoNumber true, DBAccessibleFromOPCUA true, DBAccessibleFromWebserver true, IsOnlyStoredInLoadMemory false, IsRetainMemResEnabled false, IsWriteProtectedInAS false, MemoryReserve 100
   VAR
      Work { ExternalAccessible := 'False'; ExternalVisible := 'False'; ExternalWritable := 'False'; S7_SetPoint := 'True'} : Array[1..2] of "FRK_SetWorkspace";
   END_VAR
BEGIN
END_DATA_BLOCK

DATA_BLOCK "FRK_SetStore"   // DB12
{ S7_Optimized_Access := 'TRUE' }
VERSION : 0.1
// stored: AutoNumber true, DBAccessibleFromOPCUA true, DBAccessibleFromWebserver true, IsOnlyStoredInLoadMemory false, IsRetainMemResEnabled false, IsWriteProtectedInAS false, MemoryReserve 100
   VAR RETAIN
      SchemaVersion { ExternalAccessible := 'False'; ExternalVisible := 'False'; ExternalWritable := 'False'} : UInt;
      Sets { ExternalAccessible := 'False'; ExternalVisible := 'False'; ExternalWritable := 'False'; S7_SetPoint := 'True'} : Array[1..2, 1..4] of "FRK_SetPayload";
   END_VAR
BEGIN
END_DATA_BLOCK

DATA_BLOCK "FRK_UnitScratch"   // DB13
{ S7_Optimized_Access := 'TRUE' }
VERSION : 0.1
// stored: AutoNumber true, DBAccessibleFromOPCUA true, DBAccessibleFromWebserver true, IsOnlyStoredInLoadMemory false, IsRetainMemResEnabled false, IsWriteProtectedInAS false, MemoryReserve 100
   VAR
      Response { ExternalAccessible := 'False'; ExternalVisible := 'False'; ExternalWritable := 'False'; S7_SetPoint := 'True'} : "ST_HmiResponse";
      EmptyDiagnostic { ExternalAccessible := 'False'; ExternalVisible := 'False'; ExternalWritable := 'False'; S7_SetPoint := 'True'} : "ST_Diagnostic";
      EmptyConfigEntry { ExternalAccessible := 'False'; ExternalVisible := 'False'; ExternalWritable := 'False'; S7_SetPoint := 'True'} : "ST_ConfigEntry";
      EmptyEvent { ExternalAccessible := 'False'; ExternalVisible := 'False'; ExternalWritable := 'False'; S7_SetPoint := 'True'} : "ST_AlarmEvent";
   END_VAR
BEGIN
END_DATA_BLOCK

DATA_BLOCK "GDB_AccessPersistTest"   // DB14
{ S7_Optimized_Access := 'TRUE' }
VERSION : 0.1
// stored: AutoNumber true, DBAccessibleFromOPCUA true, DBAccessibleFromWebserver true, IsOnlyStoredInLoadMemory false, IsRetainMemResEnabled false, IsWriteProtectedInAS false, MemoryReserve 100
   VAR
      Operation : Int;
      Value : DInt;
      Gate : Int;
      RotateOnLogin : Bool;
      Root : String[32];
      Applied { ExternalWritable := 'False'} : Bool;
      UsersReady { ExternalWritable := 'False'} : Bool;
      UsersLost { ExternalWritable := 'False'} : Bool;
      UserGeneration { ExternalWritable := 'False'} : UDInt;
      StartupCount { ExternalWritable := 'False'} : UDInt;
      CrcWitness { ExternalWritable := 'False'} : DWord;
      Record { ExternalAccessible := 'False'; ExternalVisible := 'False'; ExternalWritable := 'False'; S7_SetPoint := 'True'} : "ST_UserRecord";
      PolicySlot { ExternalAccessible := 'False'; ExternalVisible := 'False'; ExternalWritable := 'False'} : Int;
   END_VAR
   VAR RETAIN
      ProvisionCount { ExternalWritable := 'False'} : UDInt;
   END_VAR
BEGIN
END_DATA_BLOCK

DATA_BLOCK "GDB_AccessTest"   // DB15
{ S7_Optimized_Access := 'TRUE' }
VERSION : 0.1
// stored: AutoNumber true, DBAccessibleFromOPCUA true, DBAccessibleFromWebserver true, IsOnlyStoredInLoadMemory false, IsRetainMemResEnabled false, IsWriteProtectedInAS false, MemoryReserve 100
   VAR
      ProviderOff : Bool;
      CancelOnLogin : Bool;
      SupersedeOnLogin : Bool;
      InterruptedBusy { ExternalWritable := 'False'} : Bool;
      SupersededSequence { ExternalWritable := 'False'} : UDInt;
      InterruptRequest { ExternalAccessible := 'False'; ExternalVisible := 'False'; ExternalWritable := 'False'; S7_SetPoint := 'True'} : "ST_HmiRequest";
      HashData { ExternalAccessible := 'False'; ExternalVisible := 'False'; ExternalWritable := 'False'} : Array[0..47] of Byte;
      Hash0 { ExternalWritable := 'False'} : Array[0..31] of Byte;
      Hash1 { ExternalWritable := 'False'} : Array[0..31] of Byte;
      Hash2 { ExternalWritable := 'False'} : Array[0..31] of Byte;
      Hash3 { ExternalWritable := 'False'} : Array[0..31] of Byte;
      HashOk { ExternalWritable := 'False'} : Bool;
   END_VAR
BEGIN
END_DATA_BLOCK

DATA_BLOCK "GDB_ConfigSetTest"   // DB16
{ S7_Optimized_Access := 'TRUE' }
VERSION : 0.1
// stored: AutoNumber true, DBAccessibleFromOPCUA true, DBAccessibleFromWebserver true, IsOnlyStoredInLoadMemory false, IsRetainMemResEnabled false, IsWriteProtectedInAS false, MemoryReserve 100
   VAR
      Corrupt : Bool;
      SetName : String[80];
      Field : Int;
      Text : String[80];
      Slot { ExternalWritable := 'False'} : Int;
      RecordScope { ExternalWritable := 'False'} : String[80];
      RecordKey { ExternalWritable := 'False'} : String[160];
   END_VAR
BEGIN
END_DATA_BLOCK

DATA_BLOCK "GDB_ConfigTest"   // DB17
{ S7_Optimized_Access := 'TRUE' }
VERSION : 0.1
// stored: AutoNumber true, DBAccessibleFromOPCUA true, DBAccessibleFromWebserver true, IsOnlyStoredInLoadMemory false, IsRetainMemResEnabled false, IsWriteProtectedInAS false, MemoryReserve 100
   VAR
      Unavailable : Bool;
      CorruptPulse : Bool;
      CorruptScope : String[80];
      CorruptKey : String[160];
      CorruptModel : String[64];
      CorruptText : String[80];
      CorruptSchema : UInt;
      CorruptSlot { ExternalWritable := 'False'} : Int;
      ConfiguredPulse : Bool;
   END_VAR
   VAR RETAIN
      BlockRestore : Bool;
   END_VAR
BEGIN
END_DATA_BLOCK

DATA_BLOCK "GDB_DecisionTest"   // DB25
{ S7_Optimized_Access := 'TRUE' }
VERSION : 0.1
// Deterministic service integration checks, independent of physical press I/O.
// stored: AutoNumber true, DBAccessibleFromOPCUA true, DBAccessibleFromWebserver true, IsOnlyStoredInLoadMemory false, IsRetainMemResEnabled false, IsWriteProtectedInAS false, MemoryReserve 100
   VAR
      Done : Bool;
      Passed : Int;
      Total : Int;
      Checks : Array[1..28] of Bool;
      EmptyHmiRequest { S7_SetPoint := 'True'} : "ST_HmiRequest";
      EmptyHmiResponse { S7_SetPoint := 'True'} : "ST_HmiResponse";
      EmptyReport { S7_SetPoint := 'True'} : "ST_ReleaseReport";
      WorkRequest { ExternalAccessible := 'False'; ExternalVisible := 'False'; ExternalWritable := 'False'; S7_SetPoint := 'True'} : "ST_DecisionRequest";
      WorkPublished { ExternalAccessible := 'False'; ExternalVisible := 'False'; ExternalWritable := 'False'; S7_SetPoint := 'True'} : "ST_DecisionRequest";
      WorkReport { ExternalAccessible := 'False'; ExternalVisible := 'False'; ExternalWritable := 'False'; S7_SetPoint := 'True'} : "ST_ReleaseReport";
      WorkTestCore { ExternalAccessible := 'False'; ExternalVisible := 'False'; ExternalWritable := 'False'; S7_SetPoint := 'True'} : "FRK_Core";
      WorkTestUnit { ExternalAccessible := 'False'; ExternalVisible := 'False'; ExternalWritable := 'False'; S7_SetPoint := 'True'} : "FRK_Unit";
      WorkTestAccess { ExternalAccessible := 'False'; ExternalVisible := 'False'; ExternalWritable := 'False'; S7_SetPoint := 'True'} : "FRK_Access";
      WorkHmiRequest { ExternalAccessible := 'False'; ExternalVisible := 'False'; ExternalWritable := 'False'; S7_SetPoint := 'True'} : "ST_HmiRequest";
      WorkHmiResponse { ExternalAccessible := 'False'; ExternalVisible := 'False'; ExternalWritable := 'False'; S7_SetPoint := 'True'} : "ST_HmiResponse";
      Log { ExternalAccessible := 'False'; ExternalVisible := 'False'; ExternalWritable := 'False'; S7_SetPoint := 'True'} : "FRK_AlarmLog";
   END_VAR
BEGIN
END_DATA_BLOCK

DATA_BLOCK "GDB_FraktalHal"   // DB22
{ S7_Optimized_Access := 'TRUE' }
VERSION : 0.1
// stored: AutoNumber true, DBAccessibleFromOPCUA true, DBAccessibleFromWebserver true, IsOnlyStoredInLoadMemory false, IsRetainMemResEnabled false, IsWriteProtectedInAS false, MemoryReserve 100
   VAR
      Data { ExternalAccessible := 'False'; ExternalVisible := 'False'; ExternalWritable := 'False'; S7_SetPoint := 'True'} : "ST_FraktalHal";
   END_VAR
BEGIN
END_DATA_BLOCK

DATA_BLOCK "GDB_ManifestTest"   // DB18
{ S7_Optimized_Access := 'TRUE' }
VERSION : 0.1
// stored: AutoNumber true, DBAccessibleFromOPCUA true, DBAccessibleFromWebserver true, IsOnlyStoredInLoadMemory false, IsRetainMemResEnabled false, IsWriteProtectedInAS false, MemoryReserve 100
   VAR
      ReadLock : Bool;
   END_VAR
BEGIN
END_DATA_BLOCK

DATA_BLOCK "GDB_RoutingTest"   // DB19
{ S7_Optimized_Access := 'TRUE' }
VERSION : 0.1
// stored: AutoNumber true, DBAccessibleFromOPCUA true, DBAccessibleFromWebserver true, IsOnlyStoredInLoadMemory false, IsRetainMemResEnabled false, IsWriteProtectedInAS false, MemoryReserve 100
   VAR
      PermitOne : Bool;
      PermitTwo : Bool;
      NestedFinish : Bool;
      InnerFinish : Bool;
      NestedAccessLock : Bool;
      RootManualPermit : Bool;
      ManualAccessLock : Bool;
      LocalPulse : Bool;
      LocalKind : DInt;
      LocalValue : DInt;
      LocalAccepted { ExternalWritable := 'False'} : Bool;
      LocalFirstKind { ExternalWritable := 'False'} : DInt;
      LocalRequest { ExternalAccessible := 'False'; ExternalVisible := 'False'; ExternalWritable := 'False'; S7_SetPoint := 'True'} : "ST_HmiRequest";
      ManExecute { ExternalWritable := 'False'} : Bool;
      ManStarts { ExternalWritable := 'False'} : DInt;
   END_VAR
BEGIN
END_DATA_BLOCK

DATA_BLOCK "GDB_StateAlarmTest"   // DB20
{ S7_Optimized_Access := 'TRUE' }
VERSION : 0.1
// stored: AutoNumber true, DBAccessibleFromOPCUA true, DBAccessibleFromWebserver true, IsOnlyStoredInLoadMemory false, IsRetainMemResEnabled false, IsWriteProtectedInAS false, MemoryReserve 100
   VAR
      ClearLog : Bool;
      RaisePulse : Bool;
      GonePulse : Bool;
      FillPulse : Bool;
      CauseLive : Bool;
      PublishState : Bool;
      StateValue : Bool;
      Position : DInt;
      StateIndex : Int;
      ResetClass : DInt;
      FillCount : Int;
      Diag { S7_SetPoint := 'True'} : "ST_Diagnostic";
      Slot { ExternalWritable := 'False'} : Int;
      GoneAccepted { ExternalWritable := 'False'} : Bool;
      SinkCome { ExternalWritable := 'False'} : UDInt;
      SinkClose { ExternalWritable := 'False'} : UDInt;
      SinkLast { ExternalWritable := 'False'; S7_SetPoint := 'True'} : "ST_AlarmEvent";
      NativeFaultSlot { ExternalWritable := 'False'} : Int;
      StandaloneCount { ExternalWritable := 'False'} : Int;
      StandaloneReturn { ExternalWritable := 'False'} : Bool;
      StandaloneFlags { ExternalWritable := 'False'; S7_SetPoint := 'True'} : Array[1..12] of "ST_StateFlag";
      CauseSlot { ExternalAccessible := 'False'; ExternalVisible := 'False'; ExternalWritable := 'False'} : Int;
      Touched { ExternalAccessible := 'False'; ExternalVisible := 'False'; ExternalWritable := 'False'} : Array[1..12] of Bool;
   END_VAR
BEGIN
END_DATA_BLOCK

DATA_BLOCK "GDB_UnitTest"   // DB21
{ S7_Optimized_Access := 'TRUE' }
VERSION : 0.1
// stored: AutoNumber true, DBAccessibleFromOPCUA true, DBAccessibleFromWebserver true, IsOnlyStoredInLoadMemory false, IsRetainMemResEnabled false, IsWriteProtectedInAS false, MemoryReserve 100
   VAR
      FinishCycle : Bool;
      Permit : Bool;
      FaultRoot : Bool;
      ExitHold : Bool;
      LockStart : Bool;
      IssueChild : Bool;
      ChildCommand : DInt;
      Verdict : DInt;
      Reason : DInt;
      CarrierControl : DInt;
      Scans { ExternalWritable := 'False'} : UDInt;
      Restarts { ExternalWritable := 'False'} : UDInt;
      ChildExecute { ExternalWritable := 'False'} : Bool;
      ChildState { ExternalWritable := 'False'} : DInt;
      CarrierWrites { ExternalWritable := 'False'} : UDInt;
      CarrierSerial { ExternalWritable := 'False'} : UDInt;
      WrittenUid { ExternalWritable := 'False'} : String[64];
      WrittenVerdict { ExternalWritable := 'False'} : DInt;
      LastEvent { ExternalWritable := 'False'} : DInt;
      SecretCleared { ExternalWritable := 'False'} : Bool;
      SnapshotSecretCleared { ExternalWritable := 'False'} : Bool;
      BootStamp { ExternalWritable := 'False'} : LDT;
   END_VAR
BEGIN
END_DATA_BLOCK

ORGANIZATION_BLOCK "Main"   // OB1, SCL, ProgramCycle
TITLE = "Main Program Sweep (Cycle)"
{ S7_Optimized_Access := 'TRUE' }
VERSION : 0.1
// stored: AutoNumber true, IsIECCheckEnabled false, SetENOAutomatically false
   VAR_INPUT
      Initial_Call : Bool;   // Initial call of this OB
      Remanence : Bool;   // =True, if remanent data are available
   END_VAR
BEGIN

   "F_ConfigBenchPrepare"(Startup := #Initial_Call);
   "GDB_FraktalMain"(Startup := #Initial_Call);
   "F_ConfigBenchObserve"(Startup := #Initial_Call);
   "F_DecisionBench"();
END_ORGANIZATION_BLOCK

FUNCTION_BLOCK "FB_FraktalMain"   // FB6, SCL
{ S7_Optimized_Access := 'TRUE' }
VERSION : 0.1
// stored: AutoNumber true, IsIECCheckEnabled false, IsRetainMemResEnabled false, MemoryReserve 100, SetENOAutomatically false, UDAEnableTagReadback false
   VAR_INPUT
      Startup { ExternalAccessible := 'False'; ExternalVisible := 'False'; ExternalWritable := 'False'} : Bool;
   END_VAR
BEGIN

   IF #Startup THEN
       "FRK_Registry".Count := 0;
       "FRK_Registry".Fault := FALSE;
   END_IF;
   "FRK_ClockTick"();
   "FRK_AccessStoreBoot"(Startup := #Startup);
   "FRK_ConfigBoot"(Startup := #Startup);
   "FRK_SetBoot"(Startup := #Startup);
   "StationA"(ParentIndex := 0,
              Startup := #Startup,
              Hal := "GDB_FraktalHal".Data.StationA);
   "StationB"(ParentIndex := 0,
              Startup := #Startup,
              Hal := "GDB_FraktalHal".Data.StationB);
END_FUNCTION_BLOCK

FUNCTION_BLOCK "FB_DeclarationUnit"   // FB5, SCL
{ S7_Optimized_Access := 'TRUE' }
VERSION : 0.1
// Generated frame v0.11; change the declaration, then regenerate.
// stored: AutoNumber true, IsIECCheckEnabled false, IsRetainMemResEnabled false, MemoryReserve 100, SetENOAutomatically false, UDAEnableTagReadback false
   VAR_INPUT
      Execute { ExternalWritable := 'False'} : Bool;
      Abort { ExternalWritable := 'False'} : Bool;
      Command { ExternalWritable := 'False'} : DInt;
      ParCmd { ExternalWritable := 'False'} : "ST_DeclarationParCmd";
      ParentIndex { ExternalAccessible := 'False'; ExternalVisible := 'False'; ExternalWritable := 'False'} : DInt;
      Startup { ExternalAccessible := 'False'; ExternalVisible := 'False'; ExternalWritable := 'False'} : Bool;
   END_VAR
   VAR_OUTPUT
      Busy { ExternalWritable := 'False'} : Bool;
      Done { ExternalWritable := 'False'} : Bool;
      Error { ExternalWritable := 'False'} : Bool;
      Aborted { ExternalWritable := 'False'} : Bool;
      Held { ExternalWritable := 'False'} : Bool;
      ErrorID { ExternalWritable := 'False'} : DWord;
      Timing { ExternalWritable := 'False'} : "ST_ModuleTiming";
      OutCmd { ExternalWritable := 'False'} : "ST_DeclarationOutCmd";
      OutImm { ExternalWritable := 'False'} : "ST_UnitProbeImm";
   END_VAR
   VAR_IN_OUT
      Hal : "ST_DeclarationUnitHal";
   END_VAR
   VAR
      Status { ExternalWritable := 'False'; S7_SetPoint := 'True'} : "ST_ModuleStatus";
      Core { ExternalAccessible := 'False'; ExternalVisible := 'False'; ExternalWritable := 'False'; S7_SetPoint := 'True'} : "FRK_Core";
      ParCfg { ExternalWritable := 'False'; S7_SetPoint := 'True'} : "ST_DeclarationParCfg";
      LatchedParCmd { ExternalAccessible := 'False'; ExternalVisible := 'False'; ExternalWritable := 'False'; S7_SetPoint := 'True'} : "ST_DeclarationParCmd";
      StateFlags { ExternalWritable := 'False'; S7_SetPoint := 'True'} : Array[1..12] of "ST_StateFlag";
      StateFlagCount { ExternalWritable := 'False'} : Int;
      StateTouched { ExternalAccessible := 'False'; ExternalVisible := 'False'; ExternalWritable := 'False'} : Array[1..12] of Bool;
      Device { ExternalAccessible := 'False'; ExternalVisible := 'False'; ExternalWritable := 'False'; S7_SetPoint := 'True'} : "ST_UnitProbeDevice";
      StationCfg { ExternalWritable := 'False'; S7_SetPoint := 'True'} : "ST_UnitProbeStationCfg";
      ConfigStageParCfg { ExternalAccessible := 'False'; ExternalVisible := 'False'; ExternalWritable := 'False'; S7_SetPoint := 'True'} : "ST_DeclarationParCfg";
      ConfigDefaultParCfg { ExternalAccessible := 'False'; ExternalVisible := 'False'; ExternalWritable := 'False'; S7_SetPoint := 'True'} : "ST_DeclarationParCfg";
      ConfigStageStationCfg { ExternalAccessible := 'False'; ExternalVisible := 'False'; ExternalWritable := 'False'; S7_SetPoint := 'True'} : "ST_UnitProbeStationCfg";
      ConfigDefaultStationCfg { ExternalAccessible := 'False'; ExternalVisible := 'False'; ExternalWritable := 'False'; S7_SetPoint := 'True'} : "ST_UnitProbeStationCfg";
      ConfigStaged { ExternalAccessible := 'False'; ExternalVisible := 'False'; ExternalWritable := 'False'} : Bool;
      ConfigPersist { ExternalWritable := 'False'; S7_SetPoint := 'True'} : "ST_ConfigPersistStatus";
      ModelId { ExternalWritable := 'False'; S7_SetPoint := 'True'} : "ST_ModelId";
      AvailableModelCount { ExternalWritable := 'False'} : Int;
      AvailableModels { ExternalWritable := 'False'; S7_SetPoint := 'True'} : Array[1..2] of "ST_ModelId";
      ConfigSets { ExternalWritable := 'False'; S7_SetPoint := 'True'} : Array[1..4] of "ST_ConfigSetInfo";
      ConfigSetCount { ExternalWritable := 'False'} : Int;
      ConfigSetDocument { ExternalWritable := 'False'} : WString[480];
      ConfigSetDocumentLine { ExternalWritable := 'False'} : Int;
      ConfigSetDocumentLines { ExternalWritable := 'False'} : Int;
      Unit { ExternalAccessible := 'False'; ExternalVisible := 'False'; ExternalWritable := 'False'; S7_SetPoint := 'True'} : "FRK_Unit";
      HmiRequest { S7_SetPoint := 'True'} : "ST_HmiRequest";
      ModePolicy { ExternalAccessible := 'False'; ExternalVisible := 'False'; ExternalWritable := 'False'; S7_SetPoint := 'True'} : Array[0..6] of "ST_ModePolicy";
      Access { ExternalWritable := 'False'; S7_SetPoint := 'True'} : "FRK_Access";
      HmiResponse { ExternalWritable := 'False'; S7_SetPoint := 'True'} : "ST_HmiResponse";
      ConfigRev { ExternalWritable := 'False'} : UDInt;
      ConfigCursor { ExternalAccessible := 'False'; ExternalVisible := 'False'; ExternalWritable := 'False'; S7_SetPoint := 'True'} : "FRK_ConfigCursor";
      Part { ExternalWritable := 'False'; S7_SetPoint := 'True'} : "ST_PartContext";
      Decision { ExternalWritable := 'False'; S7_SetPoint := 'True'} : "ST_DecisionRequest";
      DecisionAnswer { ExternalWritable := 'False'} : Int;
      History { ExternalWritable := 'False'; S7_SetPoint := 'True'} : Array[1..16] of "ST_Diagnostic";
      HistoryHead { ExternalWritable := 'False'} : Int;
      AlarmLog { ExternalWritable := 'False'; S7_SetPoint := 'True'} : "FRK_AlarmLog";
      ModeActivePublished { ExternalWritable := 'False'} : DInt;
      RunningPublished { ExternalWritable := 'False'} : Bool;
      StopPendingPublished { ExternalWritable := 'False'} : Bool;
      SupportedModesPublished { ExternalWritable := 'False'} : Array[0..6] of Bool;
      GoodCount { ExternalWritable := 'False'} : UDInt;
      NokCount { ExternalWritable := 'False'} : UDInt;
      ReworkCount { ExternalWritable := 'False'} : UDInt;
      NokReason { ExternalWritable := 'False'} : DInt;
      Cell { ExternalWritable := 'False'; S7_SetPoint := 'True'} : "FB_DeclarationCell";
      Satellite { ExternalWritable := 'False'; S7_SetPoint := 'True'} : "FB_SatelliteUnit";
   END_VAR
   VAR_TEMP
      InstancePath : WString[254];
      RouteMatched : Bool;
      ManualMatched : Bool;
      ConfigRootIndex : Int;
   END_VAR
   VAR CONSTANT
      EXEC_READY : DInt := 0;
      MODULE_TIER : DInt := 1;
   END_VAR
BEGIN

   // ---- GENERATED: setup
   IF #Startup OR NOT #Core.Named THEN
       #InstancePath := GetInstancePath(size := 0);
       "FRK_SetIdentity"(Core := #Core,
                         Status := #Status,
                         InstancePath := #InstancePath,
                         ModuleType := 1,
                         TypeId := 1,
                         Capabilities := DWORD#16#00000000,
                         ParentIndex := #ParentIndex,
                         TypeKey := 'Fraktal.Declaration.Unit');
   END_IF;
   IF #Startup THEN "FRK_CfgRestore_DeclarationUnit"(Core := #Core,
                                                         Status := #Status,
                                                         ParCfg := #ParCfg,
                                                         StationCfg := #StationCfg,
                                                         ConfigStageParCfg := #ConfigStageParCfg,
                                                         ConfigDefaultParCfg := #ConfigDefaultParCfg,
                                                         ConfigStageStationCfg := #ConfigStageStationCfg,
                                                         ConfigDefaultStationCfg := #ConfigDefaultStationCfg);
   END_IF;
   #ConfigRootIndex := "FRK_ConfigRoot"(RegIndex := #Core.RegIndex);
   IF #Core.ParentIndex = 0 THEN
       #AvailableModelCount := 2;
   ELSE
       #AvailableModelCount := 0;
   END_IF;
   #AvailableModels[1].ModelCode := 'MODEL_A';
   #AvailableModels[2].ModelCode := 'MODEL_B';
   "FRK_StateSweep"(Flags := #StateFlags,
                    Count := #StateFlagCount,
                    Touched := #StateTouched,
                    Startup := #Startup);
   IF #Startup OR #ConfigRev = 0 THEN
       #ConfigRev := "FRK_ConfigRevision"(Previous := #ConfigRev);
   END_IF;
   #SupportedModesPublished[0] := TRUE;
   #SupportedModesPublished[1] := TRUE;
   #SupportedModesPublished[2] := TRUE;
   #SupportedModesPublished[3] := TRUE;
   #SupportedModesPublished[4] := FALSE;
   #SupportedModesPublished[5] := FALSE;
   #SupportedModesPublished[6] := FALSE;
   "FRK_UnitPrepare"(Core := #Core,
                     Unit := #Unit,
                     Policy := #ModePolicy,
                     Request := #HmiRequest,
                     Response := #HmiResponse,
                     Startup := #Startup,
                     InitialMode := 1);
   "FRK_AlarmBegin"(AlarmLog := #AlarmLog,
                    Startup := #Startup);
   "FRK_AccessPolicyBoot"(Access := #Access,
                          Startup := #Startup,
                          Root := #Core.ParentIndex = 0,
                          Scope := #Status.Name);
   "FRK_AccessCyclic"(Access := #Access,
                      Startup := #Startup,
                      SourcePath := STRING_TO_WSTRING(#Status.Name),
                      AlarmLog := #AlarmLog,
                      Revision := #ConfigRev);
   "FRK_UnitMailbox"(Core := #Core,
                     Unit := #Unit,
                     Status := #Status,
                     Policy := #ModePolicy,
                     Access := #Access,
                     Request := #HmiRequest,
                     Response := #HmiResponse,
                     Supported := #SupportedModesPublished);
   "FRK_ConfigStatus"(RootIndex := #ConfigRootIndex,
                      Persist := #ConfigPersist,
                      AlarmLog := #AlarmLog);
   #Unit.ConfigEnabled := #Core.ParentIndex = 0;
   #Unit.ConfigSetsEnabled := TRUE AND #Core.ParentIndex = 0;
   #Unit.ModelEnabled := #AvailableModelCount > 0;
   #Unit.ConfigBlocked := #ConfigPersist.RestoreLost AND NOT #ConfigPersist.RestoreAcknowledged AND #ConfigPersist.RestorePolicy = 1;
   #Unit.ConfigBlocked := #Unit.ConfigBlocked OR #Access.PolicyLost;
   // ---- GENERATED: begin
   "FRK_Begin"(Core := #Core,
               Status := #Status,
               Execute := #Unit.RunReq,
               Abort := (#Abort OR #Unit.AbortReq),
               Command := 1);
   IF #Core.EvCommandStart THEN
       #LatchedParCmd := #ParCmd;
       CASE #Core.Command OF
           1:
               "FRK_UnitRunStart"(Core := #Core,
                                  Status := #Status,
                                  Timeout := #ParCfg.Timeout,
                                  Label := 'Run');
           ELSE
               "FRK_Start"(Core := #Core,
                           Status := #Status,
                           Supported := FALSE,
                           Timeout := T#0ms,
                           Label := '');
       END_CASE;
   END_IF;
   IF #Core.EvCommandStart THEN
       // ---- AUTHORED: CommandStart
       #Device.Received := "FRK_PartReceived"(Core := #Core, Unit := #Unit, Status := #Status, Part := #Part, AlarmLog := #AlarmLog);
       IF #Device.Received THEN
           "FRK_PartStarted"(Unit := #Unit,
                             Status := #Status,
                             Part := #Part,
                             AlarmLog := #AlarmLog);
       END_IF;
       // ---- GENERATED: reaction end
   END_IF;
   // ---- AUTHORED: cyclic management
   IF #Hal.Cell.Clamp.BackgroundFault THEN
       "FRK_Fault"(Core := #Core,
                   Status := #Status,
                   ReasonCode := 2901,
                   Description := WSTRING#'test.unit.condition');
   END_IF;
   // ---- GENERATED: end management
   "FRK_Release_DeclarationUnit"(Unit := #Unit,
                                 Hal := #Hal);
   IF #Core.RegIndex > 0 THEN
       "FRK_Registry".Rows[#Core.RegIndex].AlarmBlocking := #AlarmLog.Blocking;
   END_IF;
   #Unit.AlarmBlocking := "FRK_AlarmTreeBlocking"(Owner := #Core.RegIndex);
   "FRK_UnitConsume"(Core := #Core,
                     Unit := #Unit,
                     Status := #Status,
                     Policy := #ModePolicy,
                     Access := #Access,
                     Response := #HmiResponse,
                     Supported := #SupportedModesPublished);
   "FRK_UnitMode"(Core := #Core,
                  Unit := #Unit);
   IF #Core.EvModeExit THEN
       // ---- AUTHORED: ModeExit
       #Device.ExitCalls := #Device.ExitCalls + 1;
       IF #Hal.Cell.Clamp.ExitHold THEN
           #Core.HookResult := 1;
       ELSE
           #Core.HookResult := 0;
       END_IF;
       // ---- GENERATED: reaction end
   END_IF;
   "FRK_UnitModeResolve"(Core := #Core,
                         Unit := #Unit,
                         Status := #Status,
                         Policy := #ModePolicy,
                         Timeout := #ParCfg.Timeout);
   IF #Core.EvModeChanged THEN
       // ---- AUTHORED: ModeChanged
       #Device.Changes := #Device.Changes + 1;
       // ---- GENERATED: reaction end
   END_IF;
   "FRK_DecisionCyclic"(Owner := #Core.RegIndex,
                        Busy := #Core.Exec = 1,
                        Reset := #Startup OR #Unit.EvReset OR #Core.EvModeChanged,
                        AlarmLog := #AlarmLog);
   "FRK_UnitFollow"(Core := #Core,
                    Unit := #Unit,
                    Status := #Status,
                    Policy := #ModePolicy,
                    Access := #Access,
                    Supported := #SupportedModesPublished);
   IF #Unit.RequestPending AND (#Unit.Request.Kind = 11 OR #Unit.Request.Kind = 16) THEN
       #ManualMatched := FALSE;
       #RouteMatched := "FRK_Route_DeclarationCell"(Module := #Cell, Hal := #Hal.Cell, Request := #Unit.Request, Report := #HmiResponse.Report);
       #ManualMatched := #ManualMatched OR #RouteMatched;
       #RouteMatched := "FRK_Route_SatelliteUnit"(Module := #Satellite, Hal := #Hal.Satellite, Request := #Unit.Request, Report := #HmiResponse.Report);
       #ManualMatched := #ManualMatched OR #RouteMatched;
       IF NOT #ManualMatched THEN
           "FRK_ReleaseReason"(Report := #HmiResponse.Report,
                               Description := WSTRING#'std.error.unsupportedHmiRequest',
                               Reason := 2008,
                               Path := #Unit.Request.TargetPath,
                               Kind := 4);
       END_IF;
       #HmiResponse.Accepted := #Unit.Request.Kind = 16 OR #HmiResponse.Report.Released;
       IF #Unit.Request.Kind = 11 THEN
           IF #HmiResponse.Accepted THEN
               #HmiResponse.Diagnostic := WSTRING#'std.audit.manualCommandAccepted';
           ELSE
               #HmiResponse.Diagnostic := WSTRING#'std.audit.manualCommandRejected';
           END_IF;
       END_IF;
   END_IF;
   IF #Unit.EvReset THEN
       "FRK_AlarmOperatorReset"(AlarmLog := #AlarmLog);
   END_IF;
   IF #Unit.EvReset THEN
       // ---- AUTHORED: OperatorReset
       #Device.Resets := #Device.Resets + 1;
       // ---- GENERATED: reset reaction end
   END_IF;
   IF #Core.ReleasePending OR #Unit.ReleaseChildren THEN
       "FRK_ReleaseCommand"(Core := #Cell.Core,
                            Execute := #Cell.Execute);
       "FRK_ReleaseCommand"(Core := #Satellite.Core,
                            Execute := #Satellite.Execute);
   END_IF;
   // ---- GENERATED: child call
   #Cell(ParentIndex := #Core.RegIndex,
         Startup := #Startup,
         Hal := #Hal.Cell);
   "FRK_ManualFinish"(Core := #Cell.Core,
                      Execute := #Cell.Execute,
                      ManualOwned := #Cell.ManualOwned);
   "FRK_UnitCascade"(ParentUnit := #Unit,
                     Core := #Satellite.Core,
                     Unit := #Satellite.Unit,
                     Status := #Satellite.Status,
                     Policy := #Satellite.ModePolicy,
                     Access := #Satellite.Access,
                     Supported := #Satellite.SupportedModesPublished,
                     AlarmLog := #AlarmLog);
   // ---- GENERATED: child call
   #Satellite(ParentIndex := #Core.RegIndex,
              Startup := #Startup,
              Hal := #Hal.Satellite);
   #Unit.CascadePending := FALSE;
   "FRK_CfgOperation_DeclarationUnit"(Core := #Core, Status := #Status, ParCfg := #ParCfg, ModePolicy := #ModePolicy, Access := #Access, Unit := #Unit, HmiResponse := #HmiResponse, ConfigPersist := #ConfigPersist, ConfigCursor := #ConfigCursor, ConfigRev := #ConfigRev, ModelId := #ModelId, AvailableModelCount := #AvailableModelCount, ConfigStaged := #ConfigStaged, SupportedModesPublished := #SupportedModesPublished, StationCfg := #StationCfg, ConfigStageParCfg := #ConfigStageParCfg, ConfigDefaultParCfg := #ConfigDefaultParCfg, Cell := #Cell, Satellite := #Satellite);
   "FRK_CfgSetOperation_DeclarationUnit"(Core := #Core, Status := #Status, ParCfg := #ParCfg, ModePolicy := #ModePolicy, Access := #Access, Unit := #Unit, HmiResponse := #HmiResponse, ConfigPersist := #ConfigPersist, ConfigRev := #ConfigRev, ModelId := #ModelId, ConfigSets := #ConfigSets, ConfigSetCount := #ConfigSetCount, ConfigSetDocument := #ConfigSetDocument, ConfigSetDocumentLine := #ConfigSetDocumentLine, ConfigSetDocumentLines := #ConfigSetDocumentLines, SupportedModesPublished := #SupportedModesPublished, StationCfg := #StationCfg, ConfigStageParCfg := #ConfigStageParCfg, ConfigStageStationCfg := #ConfigStageStationCfg, Cell := #Cell, Satellite := #Satellite, Startup := #Startup);
   IF #Unit.RequestPending AND #Core.ParentIndex = 0 THEN
       "FRK_SetResult"(Request := #Unit.Request,
                       Response := #HmiResponse,
                       Persist := #ConfigPersist,
                       AlarmLog := #AlarmLog,
                       Scope := #Status.Name,
                       RootIndex := #ConfigRootIndex);
   END_IF;
   "FRK_ConfigStatus"(RootIndex := #ConfigRootIndex,
                      Persist := #ConfigPersist,
                      AlarmLog := #AlarmLog);
   "FRK_RouteAbort"(Core := #Core,
                    Abort := (#Abort OR #Unit.AbortReq));
   IF #Core.EvAbort THEN
       "FRK_PartAborted"(Core := #Core,
                         Unit := #Unit,
                         Status := #Status,
                         Part := #Part,
                         AlarmLog := #AlarmLog);
   END_IF;
   IF #Core.Dispatch AND #Core.RegIndex > 0 AND NOT "FRK_Registry".Fault THEN
       // ---- AUTHORED: dispatch
       IF #Hal.Cell.Clamp.Finish THEN
           #Device.Processed := FALSE;
           IF #Unit.CarrierIndex = 0 THEN
               #Device.Processed := TRUE;
           ELSE
               #Device.Processed := "FRK_PartProcessed"(Core := #Core, Unit := #Unit, Status := #Status, Part := #Part, AlarmLog := #AlarmLog, Verdict := #Hal.Cell.Clamp.Verdict, Reason := #Hal.Cell.Clamp.Diag.ReasonCode);
           END_IF;
           IF #Device.Processed THEN
               #Device.Cycles := #Device.Cycles + 1;
               IF #Unit.StopReq THEN
                   "FRK_Complete"(Core := #Core,
                                  Status := #Status);
               ELSE
                   #Device.Received := "FRK_PartReceived"(Core := #Core, Unit := #Unit, Status := #Status, Part := #Part, AlarmLog := #AlarmLog);
                   IF #Device.Received THEN
                       "FRK_PartStarted"(Unit := #Unit,
                                         Status := #Status,
                                         Part := #Part,
                                         AlarmLog := #AlarmLog);
                   END_IF;
               END_IF;
           END_IF;
       END_IF;
       // ---- GENERATED: end dispatch
   END_IF;
   "FRK_End"(Core := #Core,
             Status := #Status,
             Busy => #Busy,
             Done => #Done,
             Error => #Error,
             Aborted => #Aborted,
             Held => #Held,
             ErrorID => #ErrorID,
             Timing => #Timing);
   "FRK_DecisionCyclic"(Owner := #Core.RegIndex,
                        Busy := #Core.Exec = 1,
                        Reset := #Startup OR #Unit.EvReset OR #Core.EvModeChanged,
                        AlarmLog := #AlarmLog);
   "FRK_DecisionPublish"(Owner := #Core.RegIndex,
                         Decision := #Decision,
                         DecisionAnswer := #DecisionAnswer);
   IF NOT #Unit.EvReset THEN
       "FRK_AlarmCapture"(AlarmLog := #AlarmLog,
                          Core := #Core,
                          Status := #Status);
       "FRK_Capture_DeclarationCell"(Module := #Cell,
                                     AlarmLog := #AlarmLog);
       "FRK_AlarmEnd"(AlarmLog := #AlarmLog);
   END_IF;
   IF #Core.RegIndex > 0 THEN
       "FRK_Registry".Rows[#Core.RegIndex].AlarmBlocking := #AlarmLog.Blocking;
   END_IF;
   #Unit.AlarmBlocking := "FRK_AlarmTreeBlocking"(Owner := #Core.RegIndex);
   "FRK_AccessPersist"(Access := #Access,
                       Unit := #Unit,
                       Response := #HmiResponse,
                       SourcePath := STRING_TO_WSTRING(#Status.Name),
                       AlarmLog := #AlarmLog);
   IF #Core.ParentIndex = 0 AND (#Access.PolicyLost OR "FRK_AccessStorage".UsersLost) THEN
       #ConfigPersist.RestoreLost := TRUE;
       #ConfigPersist.RestoreAcknowledged := FALSE;
       IF #Access.PolicyLost THEN
           #ConfigPersist.LostPath := CONCAT(IN1 := #Status.Name, IN2 := '.AccessPolicy');
       ELSE
           #ConfigPersist.LostPath := CONCAT(IN1 := #Status.Name, IN2 := '.Access');
       END_IF;
   END_IF;
   "FRK_AccessFinish"(Access := #Access,
                      Unit := #Unit,
                      Response := #HmiResponse,
                      SourcePath := STRING_TO_WSTRING(#Status.Name),
                      AlarmLog := #AlarmLog,
                      Revision := #ConfigRev);
   "FRK_UnitFinish"(Core := #Core,
                    Unit := #Unit,
                    Response := #HmiResponse,
                    Status := #Status,
                    Part := #Part,
                    AlarmLog := #AlarmLog,
                    History := #History,
                    Head := #HistoryHead);
   #ModeActivePublished := #Unit.Mode;
   #RunningPublished := #Core.Exec = 1;
   #StopPendingPublished := #Unit.StopReq AND #Core.Exec = 1;
   #GoodCount := #Unit.Good;
   #NokCount := #Unit.Nok;
   #ReworkCount := #Unit.Rework;
   #NokReason := #Unit.NokReason;
   // ---- AUTHORED: unconditional cyclic/derived data
   #OutImm.Cycles := #Device.Cycles;
   #OutImm.ExitCalls := #Device.ExitCalls;
   #OutImm.Changes := #Device.Changes;
   #OutImm.Resets := #Device.Resets;
   #OutImm.AtHome := "FRK_State"(Idx := 1, Key := 'project.state.atHome', Ok := #Hal.Cell.Clamp.Sample = 0, Flags := #StateFlags, Count := #StateFlagCount, Touched := #StateTouched);
   // ---- GENERATED: frame end
END_FUNCTION_BLOCK

FUNCTION_BLOCK "FB_DeclarationCell"   // FB2, SCL
{ S7_Optimized_Access := 'TRUE' }
VERSION : 0.1
// Generated frame v0.11; change the declaration, then regenerate.
// stored: AutoNumber true, IsIECCheckEnabled false, IsRetainMemResEnabled false, MemoryReserve 100, SetENOAutomatically false, UDAEnableTagReadback false
   VAR_INPUT
      Execute { ExternalWritable := 'False'} : Bool;
      Abort { ExternalWritable := 'False'} : Bool;
      Command { ExternalWritable := 'False'} : DInt;
      ParCmd { ExternalWritable := 'False'} : "ST_DeclarationParCmd";
      ParentIndex { ExternalAccessible := 'False'; ExternalVisible := 'False'; ExternalWritable := 'False'} : DInt;
      Startup { ExternalAccessible := 'False'; ExternalVisible := 'False'; ExternalWritable := 'False'} : Bool;
   END_VAR
   VAR_OUTPUT
      Busy { ExternalWritable := 'False'} : Bool;
      Done { ExternalWritable := 'False'} : Bool;
      Error { ExternalWritable := 'False'} : Bool;
      Aborted { ExternalWritable := 'False'} : Bool;
      Held { ExternalWritable := 'False'} : Bool;
      ErrorID { ExternalWritable := 'False'} : DWord;
      Timing { ExternalWritable := 'False'} : "ST_ModuleTiming";
      OutCmd { ExternalWritable := 'False'} : "ST_DeclarationOutCmd";
      OutImm { ExternalWritable := 'False'} : "ST_DeclarationOutImm";
   END_VAR
   VAR_IN_OUT
      Hal : "ST_DeclarationCellHal";
   END_VAR
   VAR
      Status { ExternalWritable := 'False'; S7_SetPoint := 'True'} : "ST_ModuleStatus";
      Core { ExternalAccessible := 'False'; ExternalVisible := 'False'; ExternalWritable := 'False'; S7_SetPoint := 'True'} : "FRK_Core";
      ParCfg { ExternalWritable := 'False'; S7_SetPoint := 'True'} : "ST_DeclarationParCfg";
      LatchedParCmd { ExternalAccessible := 'False'; ExternalVisible := 'False'; ExternalWritable := 'False'; S7_SetPoint := 'True'} : "ST_DeclarationParCmd";
      Device { ExternalAccessible := 'False'; ExternalVisible := 'False'; ExternalWritable := 'False'; S7_SetPoint := 'True'} : "ST_DeclarationOutImm";
      ConfigStageParCfg { ExternalAccessible := 'False'; ExternalVisible := 'False'; ExternalWritable := 'False'; S7_SetPoint := 'True'} : "ST_DeclarationParCfg";
      ConfigDefaultParCfg { ExternalAccessible := 'False'; ExternalVisible := 'False'; ExternalWritable := 'False'; S7_SetPoint := 'True'} : "ST_DeclarationParCfg";
      ConfigStaged { ExternalAccessible := 'False'; ExternalVisible := 'False'; ExternalWritable := 'False'} : Bool;
      Catalog { ExternalAccessible := 'False'; ExternalVisible := 'False'; ExternalWritable := 'False'; S7_SetPoint := 'True'} : Array[1..12] of "ST_CommandInfo";
      CatalogCount { ExternalAccessible := 'False'; ExternalVisible := 'False'; ExternalWritable := 'False'} : Int;
      ManConditions { ExternalAccessible := 'False'; ExternalVisible := 'False'; ExternalWritable := 'False'; S7_SetPoint := 'True'} : Array[1..16] of "FRK_ManualConditionRow";
      ManualOwned { ExternalAccessible := 'False'; ExternalVisible := 'False'; ExternalWritable := 'False'} : Bool;
      Clamp { ExternalWritable := 'False'; S7_SetPoint := 'True'} : "FB_DeclarationCylinder";
      Gate { ExternalWritable := 'False'; S7_SetPoint := 'True'} : "FB_DeclarationCylinder";
   END_VAR
   VAR_TEMP
      InstancePath : WString[254];
   END_VAR
   VAR CONSTANT
      EXEC_READY : DInt := 0;
      MODULE_TIER : DInt := 2;
   END_VAR
BEGIN

   // ---- GENERATED: setup
   IF #Startup OR NOT #Core.Named THEN
       #InstancePath := GetInstancePath(size := 0);
       "FRK_SetIdentity"(Core := #Core,
                         Status := #Status,
                         InstancePath := #InstancePath,
                         ModuleType := 2,
                         TypeId := 2,
                         Capabilities := DWORD#16#00000000,
                         ParentIndex := #ParentIndex,
                         TypeKey := 'Fraktal.Declaration.Cell');
       #CatalogCount := 7;
       #Catalog[1].Value := 1;
       #Catalog[1].Label := 'Finish';
       #Catalog[1].Style := 0;
       #Catalog[2].Value := 2;
       #Catalog[2].Label := 'Wait';
       #Catalog[2].Style := 0;
       #Catalog[3].Value := 3;
       #Catalog[3].Label := 'Hold';
       #Catalog[3].Style := 0;
       #Catalog[4].Value := 4;
       #Catalog[4].Label := 'Fault';
       #Catalog[4].Style := 0;
       #Catalog[5].Value := 5;
       #Catalog[5].Label := 'Pending';
       #Catalog[5].Style := 0;
       #Catalog[6].Value := 6;
       #Catalog[6].Label := 'Instant';
       #Catalog[6].Style := 0;
       #Catalog[7].Value := 7;
       #Catalog[7].Label := 'Adopt';
       #Catalog[7].Style := 0;
   END_IF;
   IF #Startup THEN "FRK_CfgRestore_DeclarationCell"(Core := #Core,
                                                         Status := #Status,
                                                         ParCfg := #ParCfg,
                                                         ConfigStageParCfg := #ConfigStageParCfg,
                                                         ConfigDefaultParCfg := #ConfigDefaultParCfg);
   END_IF;
   // ---- GENERATED: begin
   "FRK_Begin"(Core := #Core,
               Status := #Status,
               Execute := #Execute,
               Abort := #Abort,
               Command := #Command);
   IF #Core.EvInit THEN
       // ---- AUTHORED: Init
       #Device.InitCount := #Device.InitCount + 1;
       // ---- GENERATED: reaction end
   END_IF;
   IF #Core.EvCommandStart THEN
       #LatchedParCmd := #ParCmd;
       CASE #Core.Command OF
           1:
               "FRK_Start"(Core := #Core,
                           Status := #Status,
                           Supported := TRUE,
                           Timeout := #ParCfg.Timeout,
                           Label := 'Finish');
           2:
               "FRK_Start"(Core := #Core,
                           Status := #Status,
                           Supported := TRUE,
                           Timeout := #ParCfg.Timeout,
                           Label := 'Wait');
           3:
               "FRK_Start"(Core := #Core,
                           Status := #Status,
                           Supported := TRUE,
                           Timeout := #ParCfg.Timeout,
                           Label := 'Hold');
           4:
               "FRK_Start"(Core := #Core,
                           Status := #Status,
                           Supported := TRUE,
                           Timeout := #ParCfg.Timeout,
                           Label := 'Fault');
           5:
               "FRK_Start"(Core := #Core,
                           Status := #Status,
                           Supported := TRUE,
                           Timeout := #ParCfg.Timeout,
                           Label := 'Pending');
           6:
               "FRK_Start"(Core := #Core,
                           Status := #Status,
                           Supported := TRUE,
                           Timeout := #ParCfg.Timeout,
                           Label := 'Instant');
           7:
               "FRK_Start"(Core := #Core,
                           Status := #Status,
                           Supported := TRUE,
                           Timeout := #ParCfg.Timeout,
                           Label := 'Adopt');
           ELSE
               "FRK_Start"(Core := #Core,
                           Status := #Status,
                           Supported := FALSE,
                           Timeout := T#0ms,
                           Label := '');
       END_CASE;
   END_IF;
   IF #Core.EvCommandStart THEN
       // ---- AUTHORED: CommandStart
       #Device.StartCount := #Device.StartCount + 1;
       #Device.Ordered := #Device.InitCount = 1;
       // ---- GENERATED: reaction end
   END_IF;
   IF #Core.ReleasePending THEN
       "FRK_ReleaseCommand"(Core := #Clamp.Core,
                            Execute := #Clamp.Execute);
       "FRK_ReleaseCommand"(Core := #Gate.Core,
                            Execute := #Gate.Execute);
   END_IF;
   // ---- GENERATED: child call
   #Clamp(ParentIndex := #Core.RegIndex,
          Startup := #Startup,
          Hal := #Hal.Clamp);
   "FRK_ManualFinish"(Core := #Clamp.Core,
                      Execute := #Clamp.Execute,
                      ManualOwned := #Clamp.ManualOwned);
   // ---- GENERATED: child call
   #Gate(ParentIndex := #Core.RegIndex,
         Startup := #Startup,
         Hal := #Hal.Gate);
   "FRK_ManualFinish"(Core := #Gate.Core,
                      Execute := #Gate.Execute,
                      ManualOwned := #Gate.ManualOwned);
   "FRK_RouteAbort"(Core := #Core,
                    Abort := #Abort);
   "FRK_End"(Core := #Core,
             Status := #Status,
             Busy => #Busy,
             Done => #Done,
             Error => #Error,
             Aborted => #Aborted,
             Held => #Held,
             ErrorID => #ErrorID,
             Timing => #Timing);
   // ---- AUTHORED: unconditional cyclic/derived data
   #Device.Sample := #Device.Sample + 1;
   #OutImm := #Device;
   // ---- GENERATED: frame end
END_FUNCTION_BLOCK

FUNCTION_BLOCK "FB_DeclarationCylinder"   // FB1, SCL
{ S7_Optimized_Access := 'TRUE' }
VERSION : 0.1
// Generated frame v0.11; change the declaration, then regenerate.
// stored: AutoNumber true, IsIECCheckEnabled false, IsRetainMemResEnabled false, MemoryReserve 100, SetENOAutomatically false, UDAEnableTagReadback false
   VAR_INPUT
      Execute { ExternalWritable := 'False'} : Bool;
      Abort { ExternalWritable := 'False'} : Bool;
      Command { ExternalWritable := 'False'} : DInt;
      ParCmd { ExternalWritable := 'False'} : "ST_DeclarationParCmd";
      ParentIndex { ExternalAccessible := 'False'; ExternalVisible := 'False'; ExternalWritable := 'False'} : DInt;
      Startup { ExternalAccessible := 'False'; ExternalVisible := 'False'; ExternalWritable := 'False'} : Bool;
   END_VAR
   VAR_OUTPUT
      Busy { ExternalWritable := 'False'} : Bool;
      Done { ExternalWritable := 'False'} : Bool;
      Error { ExternalWritable := 'False'} : Bool;
      Aborted { ExternalWritable := 'False'} : Bool;
      Held { ExternalWritable := 'False'} : Bool;
      ErrorID { ExternalWritable := 'False'} : DWord;
      Timing { ExternalWritable := 'False'} : "ST_ModuleTiming";
      OutCmd { ExternalWritable := 'False'} : "ST_DeclarationOutCmd";
      OutImm { ExternalWritable := 'False'} : "ST_DeclarationOutImm";
   END_VAR
   VAR_IN_OUT
      Hal : "ST_DeclarationLeafHal";
   END_VAR
   VAR
      Status { ExternalWritable := 'False'; S7_SetPoint := 'True'} : "ST_ModuleStatus";
      Core { ExternalAccessible := 'False'; ExternalVisible := 'False'; ExternalWritable := 'False'; S7_SetPoint := 'True'} : "FRK_Core";
      ParCfg { ExternalWritable := 'False'; S7_SetPoint := 'True'} : "ST_DeclarationParCfg";
      LatchedParCmd { ExternalAccessible := 'False'; ExternalVisible := 'False'; ExternalWritable := 'False'; S7_SetPoint := 'True'} : "ST_DeclarationParCmd";
      Device { ExternalAccessible := 'False'; ExternalVisible := 'False'; ExternalWritable := 'False'; S7_SetPoint := 'True'} : "ST_DeclarationOutImm";
      ConfigStageParCfg { ExternalAccessible := 'False'; ExternalVisible := 'False'; ExternalWritable := 'False'; S7_SetPoint := 'True'} : "ST_DeclarationParCfg";
      ConfigDefaultParCfg { ExternalAccessible := 'False'; ExternalVisible := 'False'; ExternalWritable := 'False'; S7_SetPoint := 'True'} : "ST_DeclarationParCfg";
      ConfigStaged { ExternalAccessible := 'False'; ExternalVisible := 'False'; ExternalWritable := 'False'} : Bool;
      Catalog { ExternalAccessible := 'False'; ExternalVisible := 'False'; ExternalWritable := 'False'; S7_SetPoint := 'True'} : Array[1..12] of "ST_CommandInfo";
      CatalogCount { ExternalAccessible := 'False'; ExternalVisible := 'False'; ExternalWritable := 'False'} : Int;
      ManConditions { ExternalAccessible := 'False'; ExternalVisible := 'False'; ExternalWritable := 'False'; S7_SetPoint := 'True'} : Array[1..16] of "FRK_ManualConditionRow";
      ManualOwned { ExternalAccessible := 'False'; ExternalVisible := 'False'; ExternalWritable := 'False'} : Bool;
   END_VAR
   VAR_TEMP
      InstancePath : WString[254];
   END_VAR
   VAR CONSTANT
      EXEC_READY : DInt := 0;
      MODULE_TIER : DInt := 3;
   END_VAR
BEGIN

   // ---- GENERATED: setup
   IF #Startup OR NOT #Core.Named THEN
       #InstancePath := GetInstancePath(size := 0);
       "FRK_SetIdentity"(Core := #Core,
                         Status := #Status,
                         InstancePath := #InstancePath,
                         ModuleType := 3,
                         TypeId := 3,
                         Capabilities := DWORD#16#00000000,
                         ParentIndex := #ParentIndex,
                         TypeKey := 'Fraktal.Declaration.Cylinder');
       #CatalogCount := 7;
       #Catalog[1].Value := 1;
       #Catalog[1].Label := 'Finish';
       #Catalog[1].Style := 0;
       #Catalog[2].Value := 2;
       #Catalog[2].Label := 'Wait';
       #Catalog[2].Style := 0;
       #Catalog[3].Value := 3;
       #Catalog[3].Label := 'Hold';
       #Catalog[3].Style := 0;
       #Catalog[4].Value := 4;
       #Catalog[4].Label := 'Fault';
       #Catalog[4].Style := 0;
       #Catalog[5].Value := 5;
       #Catalog[5].Label := 'Pending';
       #Catalog[5].Style := 0;
       #Catalog[6].Value := 6;
       #Catalog[6].Label := 'Instant';
       #Catalog[6].Style := 0;
       #Catalog[7].Value := 7;
       #Catalog[7].Label := 'Adopt';
       #Catalog[7].Style := 0;
   END_IF;
   IF #Startup THEN "FRK_CfgRestore_DeclarationCylinder"(Core := #Core,
                                                             Status := #Status,
                                                             ParCfg := #ParCfg,
                                                             ConfigStageParCfg := #ConfigStageParCfg,
                                                             ConfigDefaultParCfg := #ConfigDefaultParCfg);
   END_IF;
   // ---- GENERATED: begin
   "FRK_Begin"(Core := #Core,
               Status := #Status,
               Execute := #Execute,
               Abort := #Abort,
               Command := #Command);
   IF #Core.EvInit THEN
       // ---- AUTHORED: Init
       #Device.InitCount := #Device.InitCount + 1;
       // ---- GENERATED: reaction end
   END_IF;
   IF #Core.EvCommandStart THEN
       #LatchedParCmd := #ParCmd;
       CASE #Core.Command OF
           1:
               "FRK_Start"(Core := #Core,
                           Status := #Status,
                           Supported := TRUE,
                           Timeout := #ParCfg.Timeout,
                           Label := 'Finish');
           2:
               "FRK_Start"(Core := #Core,
                           Status := #Status,
                           Supported := TRUE,
                           Timeout := #ParCfg.Timeout,
                           Label := 'Wait');
           3:
               "FRK_Start"(Core := #Core,
                           Status := #Status,
                           Supported := TRUE,
                           Timeout := #ParCfg.Timeout,
                           Label := 'Hold');
           4:
               "FRK_Start"(Core := #Core,
                           Status := #Status,
                           Supported := TRUE,
                           Timeout := #ParCfg.Timeout,
                           Label := 'Fault');
           5:
               "FRK_Start"(Core := #Core,
                           Status := #Status,
                           Supported := TRUE,
                           Timeout := #ParCfg.Timeout,
                           Label := 'Pending');
           6:
               "FRK_Start"(Core := #Core,
                           Status := #Status,
                           Supported := TRUE,
                           Timeout := #ParCfg.Timeout,
                           Label := 'Instant');
           7:
               "FRK_Start"(Core := #Core,
                           Status := #Status,
                           Supported := TRUE,
                           Timeout := #ParCfg.Timeout,
                           Label := 'Adopt');
           ELSE
               "FRK_Start"(Core := #Core,
                           Status := #Status,
                           Supported := FALSE,
                           Timeout := T#0ms,
                           Label := '');
       END_CASE;
   END_IF;
   IF #Core.EvCommandStart THEN
       // ---- AUTHORED: CommandStart
       #Device.StartCount := #Device.StartCount + 1;
       #Device.Ordered := #Device.InitCount = 1;
       // ---- GENERATED: reaction end
   END_IF;
   // ---- AUTHORED: cyclic management
   #Device.CyclicCount := #Device.CyclicCount + 1;
   IF #Hal.BackgroundFault THEN
       "FRK_Fault"(Core := #Core,
                   Status := #Status,
                   ReasonCode := 2901,
                   Description := WSTRING#'test.background');
   END_IF;
   // ---- GENERATED: end management
   "FRK_RouteAbort"(Core := #Core,
                    Abort := #Abort);
   IF #Core.EvAbort THEN
       // ---- AUTHORED: Abort
       #Device.AbortCount := #Device.AbortCount + 1;
       // ---- GENERATED: reaction end
   END_IF;
   IF #Core.EvAbortInError THEN
       // ---- AUTHORED: AbortInError
       #Device.ErrorAbortCount := #Device.ErrorAbortCount + 1;
       // ---- GENERATED: reaction end
   END_IF;
   IF #Core.Dispatch AND #Core.RegIndex > 0 AND NOT "FRK_Registry".Fault THEN
       // ---- AUTHORED: dispatch
       #Device.DispatchCount := #Device.DispatchCount + 1;
       #Device.SeenValue := #LatchedParCmd.Value;
       CASE #Core.Command OF
           1:
               IF #Hal.Finish THEN
                   #OutCmd.Result := #LatchedParCmd.Value;
                   "FRK_Complete"(Core := #Core,
                                  Status := #Status);
               END_IF;
           2:
               #Device.SeenValue := #LatchedParCmd.Value;
           3:
               IF NOT #Hal.Permit THEN
                   "FRK_Hold"(Core := #Core,
                              Status := #Status,
                              ReasonCode := 2003,
                              Description := WSTRING#'test.permit');
               ELSIF #Hal.Finish THEN
                   "FRK_Complete"(Core := #Core,
                                  Status := #Status);
               END_IF;
           4:
               "FRK_Fault"(Core := #Core,
                           Status := #Status,
                           ReasonCode := 2901,
                           Description := WSTRING#'test.first');
               "FRK_Fault"(Core := #Core,
                           Status := #Status,
                           ReasonCode := 2001,
                           Description := WSTRING#'test.second');
           5:
               "FRK_Pending"(Core := #Core,
                             Status := #Status,
                             Diag := #Hal.Diag);
               "FRK_Pending"(Core := #Core,
                             Status := #Status,
                             Diag := #Hal.LaterDiag);
           6:
               "FRK_Complete"(Core := #Core,
                              Status := #Status);
           7:
               "FRK_AdoptFault"(Core := #Core,
                                Status := #Status,
                                Diag := #Hal.Diag);
           ELSE
               "FRK_Fault"(Core := #Core,
                           Status := #Status,
                           ReasonCode := 2008,
                           Description := WSTRING#'std.error.unsupportedHmiRequest');
       END_CASE;
       // ---- GENERATED: end dispatch
   END_IF;
   "FRK_End"(Core := #Core,
             Status := #Status,
             Busy => #Busy,
             Done => #Done,
             Error => #Error,
             Aborted => #Aborted,
             Held => #Held,
             ErrorID => #ErrorID,
             Timing => #Timing);
   // ---- AUTHORED: unconditional cyclic/derived data
   #Device.Sample := #Hal.Sample;
   #Device.Output := #Core.Exec = 1 AND NOT #Core.Held AND #Hal.Permit;
   #OutImm := #Device;
   // ---- GENERATED: frame end
END_FUNCTION_BLOCK

